// TIA Portal V20 program export: 0 tag tables, 0 data types, 16 data blocks, 79 code blocks (in call order from the OBs), 59 instance data blocks

DATA_BLOCK "Control_DB"   // DB69
{ S7_Optimized_Access := 'TRUE' }
VERSION : 0.1
// stored: AutoNumber true, DBAccessibleFromOPCUA true, DBAccessibleFromWebserver true, IsOnlyStoredInLoadMemory false, IsRetainMemResEnabled false, IsWriteProtectedInAS false, MemoryReserve 100
   VAR
      Inbound_Cnv : "Inbound_Cnv_Control_UDT";
      PopUp_Cnv { S7_SetPoint := 'True'} : Array[1..4] of "PopUp_Cnv_Control";
      Outbound_Cnv { S7_SetPoint := 'True'} : "Outbound_Cnv_Control";
      ECnv_Control { S7_SetPoint := 'True'} : "ECnv_Control";
      LCnv_Control { S7_SetPoint := 'True'} : Array[1..3] of "Buffer_Cnv_Control";
      VTD_Control { S7_SetPoint := 'True'} : "VTD_Control";
      "VTD_Order Table" { S7_SetPoint := 'True'} : "WMS_OPC_UA";
      "Carrousel_Order Table" { S7_SetPoint := 'True'} : "WMS_OPC_UA";
      Shuttles_Position : Array[1..3] of Struct
         x : DInt;
         y : DInt;
         Charging : Bool;
      END_STRUCT;
      "Weighing Station" : Struct
         Start : Bool;
         Ready : Bool;
         Running : Bool;
         Done : Bool;
         Valid : Bool;
         Weight : Real;
         Error_ID : Word;
      END_STRUCT;
      "Profiling Station" : Struct
         Start : Bool;
         Ready : Bool;
         Running : Bool;
         Done : Bool;
         Valid : Bool;
         OverWidth : Bool;
         OverHeight : Bool;
         OverLength : Bool;
         Error_ID : Word;
      END_STRUCT;
      Pick_Station : Struct
         Cnv_Occupied { ExternalWritable := 'False'} : Bool;
         PushButton : Bool;
         LightGuard : Bool;
         PushButtonLight : Bool;
         Mode { ExternalWritable := 'False'} : UInt;
         Error { ExternalWritable := 'False'} : Bool;
         Warning { ExternalWritable := 'False'} : UInt;
         Enabled { ExternalWritable := 'False'} : Bool;
         Stopped { ExternalWritable := 'False'} : Bool;
         Done : Bool;
         Running { ExternalWritable := 'False'} : Bool;
         Ready_For_Task { ExternalWritable := 'False'} : Bool;
         Current_Task_Type : UInt;
         Current_Task_ID { ExternalWritable := 'False'} : UInt;
         Pallet_Type { ExternalWritable := 'False'} : UInt;
         SM_State { ExternalWritable := 'False'} : UInt;
         Motor : "Cnv_Motor";
         Instruction : "OutCnv_Instruction";
         Cnv_Errors { S7_SetPoint := 'True'} : "Cnv_Errors";
      END_STRUCT;
      InBarcode_Station : Struct
         Start : Bool;
         Ready : Bool;
         Running : Bool;
         Done : Bool;
         Valid : Bool;
         Barcode : String;
         "Reading Gate number" : String;
         "Reading Gate number OLD" : String;
         "Number of Reading Gates" : String;
         "Number of Reading Gates OLD" : String;
      END_STRUCT;
      OutBarcode_Station : Struct
         Start : Bool;
         Ready : Bool;
         Running : Bool;
         Done : Bool;
         Valid : Bool;
         Barcode : String;
         Barcode_Old : Array[1..16] of Char;
      END_STRUCT;
      VTDBarcode_Station : Struct
         Start : Bool;
         Ready : Bool;
         Running : Bool;
         Done : Bool;
         Valid : Bool;
         Barcode : String;
         Barcode_Old : String;
      END_STRUCT;
      Movement_Completed : Struct
         RTR_ITP1 : Bool;
         RTR_P1TP2 : Bool;
         RTR_P2TP3 : Bool;
         RTR_P3TP4 : Bool;
         RTR_P4TO : Bool;
         Chain_To_Chain : Bool;
         Pop4_To_Pick : Bool;
         Pick_To_Pop1 : Bool;
         WeighingStation : Bool;
      END_STRUCT;
   END_VAR
BEGIN
END_DATA_BLOCK

DATA_BLOCK "DB_SICK_AFx60_Data"   // DB120
{ S7_Optimized_Access := 'TRUE' }
VERSION : 0.1
// stored: AutoNumber true, DBAccessibleFromOPCUA true, DBAccessibleFromWebserver true, IsOnlyStoredInLoadMemory false, IsRetainMemResEnabled false, IsWriteProtectedInAS false, MemoryReserve 100
   VAR
      Data { S7_SetPoint := 'True'} : "ST_SICK_AFx60";
   END_VAR
BEGIN
END_DATA_BLOCK

DATA_BLOCK "HMI_DB"   // DB21
{ S7_Optimized_Access := 'TRUE' }
VERSION : 0.1
// stored: AutoNumber true, DBAccessibleFromOPCUA true, DBAccessibleFromWebserver true, IsOnlyStoredInLoadMemory false, IsRetainMemResEnabled false, IsWriteProtectedInAS false, MemoryReserve 100
   VAR
      Reset : Bool;
      ChargeData : Bool;
      Username : String := 'admin';
      Password : String := '12345';
      ScreenNo : UInt;
      GeneralErrors : Word;
   END_VAR
BEGIN
END_DATA_BLOCK

DATA_BLOCK "HMI_OrderTable"   // DB110
{ S7_Optimized_Access := 'TRUE' }
VERSION : 0.1
// stored: AutoNumber true, DBAccessibleFromOPCUA true, DBAccessibleFromWebserver true, IsOnlyStoredInLoadMemory false, IsRetainMemResEnabled false, IsWriteProtectedInAS false, MemoryReserve 100
   VAR
      OrderTable_1 : Array[0..9] of "OrderTable_UDT";
      OrderTable_2 : Array[0..9] of "OrderTable_UDT";
      State_1 { S7_SetPoint := 'True'} : Array[0..9] of USInt;
      State_2 { S7_SetPoint := 'True'} : Array[0..9] of USInt;
      Index_1 : Array[0..9] of Int;
      Index_2 : Array[0..9] of Int;
      ScrollUp_PB : Bool;
      ScrollDown_PB : Bool;
      PlaceOrder_PB : Bool;
      PauseOrders_PB : Bool;
      ResumeOrder_PB : Bool;
      CancelOrder_PB : Bool;
      CancelThisOrder_PB : Bool;
      StartRow : Int;
      Device : USInt;
      PlacingNewOrder : Bool;
      PopUp_ErrorWindow_Active : Bool;
      PopUp_ErrorID : UInt;
      PopUp_Index : Int;
   END_VAR
BEGIN
END_DATA_BLOCK

DATA_BLOCK "HMI_Systems"   // DB137
{ S7_Optimized_Access := 'TRUE' }
VERSION : 0.1
// stored: AutoNumber true, DBAccessibleFromOPCUA true, DBAccessibleFromWebserver true, IsOnlyStoredInLoadMemory false, IsRetainMemResEnabled false, IsWriteProtectedInAS false, MemoryReserve 100
   VAR
      SystemNo : USInt := 1;   // System Number (1 or 2)
      System { ExternalWritable := 'False'} : "System_UDT";
      CarMeasurement { ExternalWritable := 'False'} : "CarMeasurement_DB_UDT";
      EntryGate : Struct
         Sts_Opened : Bool := TRUE;
         Sts_Closed : Bool := FALSE;
         Cmd_Open : Bool := FALSE;
         Cmd_Close : Bool := FALSE;
      END_STRUCT;
      ExitGate : Struct
         Sts_Opened : Bool := TRUE;
         Sts_Closed : Bool := FALSE;
         Cmd_Open : Bool := FALSE;
         Cmd_Close : Bool := FALSE;
      END_STRUCT;
      FieldSensors : DWord := 16#04A3_7FF3;   // Field Values of Sensors
      PanelSensors : DWord := 16#04A3_7FF3;   // Sensors to show on HMI screen
      Motors : DWord := 16#0E00_6001;   // Motors to show on HMI screen
      HMI_E_Stop_System_1 : Bool := FALSE;   // HMI Emergancy Stop Push Button for System #1
      HMI_E_Stop_System_2 : Bool := FALSE;   // HMI Emergancy Stop Push Button for System #2
      HMI_E_Stop_System_3 : Bool := FALSE;   // HMI Emergancy Stop Push Button for System #2
      Virtual_Emergency_BT : Bool := false;   // HMI Emergency Stop Push Button for General system
   END_VAR
BEGIN
   System.CancelOrders := FALSE;
   System.PauseOrders := FALSE;
   System.ResumeOrders := FALSE;
   System.OrderSent := FALSE;
   System.CurrentOrder := 0;
   System.NextOrder := 1;
   System.OrderTable[0].OrderNo := 0;
   System.OrderTable[1..34].OrderNo := -1;
   System.OrderTable[35].OrderNo := 55;
   System.OrderTable[36].OrderNo := 54;
   System.OrderTable[37..38].OrderNo := 53;
   System.OrderTable[39..45].OrderNo := -1;
   System.OrderTable[46..47].OrderNo := 52;
   System.OrderTable[48..49].OrderNo := 51;
   System.OrderTable[50].OrderNo := -1;
   System.OrderTable[51].OrderNo := 50;
   System.OrderTable[52].OrderNo := 49;
   System.OrderTable[53..54].OrderNo := 48;
   System.OrderTable[55..56].OrderNo := 47;
   System.OrderTable[57..58].OrderNo := 46;
   System.OrderTable[59..60].OrderNo := 45;
   System.OrderTable[61..67].OrderNo := 44;
   System.OrderTable[68..72].OrderNo := 43;
   System.OrderTable[73..78].OrderNo := 42;
   System.OrderTable[79..80].OrderNo := 41;
   System.OrderTable[81..82].OrderNo := 40;
   System.OrderTable[83..89].OrderNo := 39;
   System.OrderTable[90..91].OrderNo := 38;
   System.OrderTable[92..96].OrderNo := 37;
   System.OrderTable[97..99].OrderNo := 36;
   System.OrderTable[0].StepNo := 0;
   System.OrderTable[1..34].StepNo := -1;
   System.OrderTable[35..36].StepNo := 1;
   System.OrderTable[37].StepNo := 2;
   System.OrderTable[38].StepNo := 1;
   System.OrderTable[39..45].StepNo := -1;
   System.OrderTable[46].StepNo := 2;
   System.OrderTable[47].StepNo := 1;
   System.OrderTable[48].StepNo := 2;
   System.OrderTable[49].StepNo := 1;
   System.OrderTable[50].StepNo := -1;
   System.OrderTable[51..52].StepNo := 1;
   System.OrderTable[53].StepNo := 2;
   System.OrderTable[54].StepNo := 1;
   System.OrderTable[55].StepNo := 2;
   System.OrderTable[56].StepNo := 1;
   System.OrderTable[57].StepNo := 2;
   System.OrderTable[58].StepNo := 1;
   System.OrderTable[59].StepNo := 2;
   System.OrderTable[60].StepNo := 1;
   System.OrderTable[61].StepNo := 7;
   System.OrderTable[62].StepNo := 6;
   System.OrderTable[63].StepNo := 5;
   System.OrderTable[64].StepNo := 4;
   System.OrderTable[65].StepNo := 3;
   System.OrderTable[66].StepNo := 2;
   System.OrderTable[67].StepNo := 1;
   System.OrderTable[68].StepNo := 5;
   System.OrderTable[69].StepNo := 4;
   System.OrderTable[70].StepNo := 3;
   System.OrderTable[71].StepNo := 2;
   System.OrderTable[72].StepNo := 1;
   System.OrderTable[73].StepNo := 6;
   System.OrderTable[74].StepNo := 5;
   System.OrderTable[75].StepNo := 4;
   System.OrderTable[76].StepNo := 3;
   System.OrderTable[77].StepNo := 2;
   System.OrderTable[78].StepNo := 1;
   System.OrderTable[79].StepNo := 2;
   System.OrderTable[80].StepNo := 1;
   System.OrderTable[81].StepNo := 2;
   System.OrderTable[82].StepNo := 1;
   System.OrderTable[83].StepNo := 7;
   System.OrderTable[84].StepNo := 6;
   System.OrderTable[85].StepNo := 5;
   System.OrderTable[86].StepNo := 4;
   System.OrderTable[87].StepNo := 3;
   System.OrderTable[88].StepNo := 2;
   System.OrderTable[89].StepNo := 1;
   System.OrderTable[90].StepNo := 2;
   System.OrderTable[91].StepNo := 1;
   System.OrderTable[92].StepNo := 5;
   System.OrderTable[93].StepNo := 4;
   System.OrderTable[94].StepNo := 3;
   System.OrderTable[95].StepNo := 2;
   System.OrderTable[96].StepNo := 1;
   System.OrderTable[97].StepNo := 6;
   System.OrderTable[98].StepNo := 5;
   System.OrderTable[99].StepNo := 4;
   System.OrderTable[0].PlaceTime := '';
   System.OrderTable[1].PlaceTime := '06/10/2022 08:58:28';
   System.OrderTable[2].PlaceTime := '06/10/2022 08:58:01';
   System.OrderTable[3].PlaceTime := '06/10/2022 08:57:38';
   System.OrderTable[4].PlaceTime := '06/10/2022 08:56:58';
   System.OrderTable[5].PlaceTime := '06/10/2022 08:46:55';
   System.OrderTable[6].PlaceTime := '06/10/2022 08:46:40';
   System.OrderTable[7].PlaceTime := '06/10/2022 08:46:00';
   System.OrderTable[8].PlaceTime := '06/10/2022 08:45:39';
   System.OrderTable[9].PlaceTime := '06/10/2022 08:45:25';
   System.OrderTable[10].PlaceTime := '06/10/2022 08:45:12';
   System.OrderTable[11].PlaceTime := '06/10/2022 08:44:47';
   System.OrderTable[12].PlaceTime := '06/10/2022 08:44:29';
   System.OrderTable[13].PlaceTime := '06/10/2022 08:44:13';
   System.OrderTable[14].PlaceTime := '06/10/2022 08:43:18';
   System.OrderTable[15].PlaceTime := '06/10/2022 08:42:58';
   System.OrderTable[16].PlaceTime := '06/10/2022 08:41:58';
   System.OrderTable[17].PlaceTime := '06/10/2022 08:41:36';
   System.OrderTable[18].PlaceTime := '06/10/2022 08:37:44';
   System.OrderTable[19].PlaceTime := '06/10/2022 08:37:27';
   System.OrderTable[20].PlaceTime := '06/10/2022 08:37:06';
   System.OrderTable[21].PlaceTime := '06/10/2022 08:35:40';
   System.OrderTable[22].PlaceTime := '06/10/2022 08:14:06';
   System.OrderTable[23].PlaceTime := '06/10/2022 08:13:36';
   System.OrderTable[24].PlaceTime := '06/10/2022 08:09:48';
   System.OrderTable[25].PlaceTime := '06/10/2022 08:09:26';
   System.OrderTable[26].PlaceTime := '06/10/2022 08:08:29';
   System.OrderTable[27].PlaceTime := '06/10/2022 08:05:42';
   System.OrderTable[28].PlaceTime := '06/10/2022 08:04:48';
   System.OrderTable[29].PlaceTime := '06/10/2022 08:03:07';
   System.OrderTable[30].PlaceTime := '06/10/2022 08:01:46';
   System.OrderTable[31].PlaceTime := '06/10/2022 08:00:57';
   System.OrderTable[32].PlaceTime := '06/10/2022 07:54:12';
   System.OrderTable[33].PlaceTime := '06/10/2022 07:53:12';
   System.OrderTable[34].PlaceTime := '06/10/2022 07:52:34';
   System.OrderTable[35].PlaceTime := '06/09/2022 15:57:28';
   System.OrderTable[36].PlaceTime := '06/09/2022 15:54:31';
   System.OrderTable[37..38].PlaceTime := '06/09/2022 15:46:22';
   System.OrderTable[39].PlaceTime := '06/09/2022 15:44:20';
   System.OrderTable[40].PlaceTime := '06/09/2022 15:44:17';
   System.OrderTable[41].PlaceTime := '06/09/2022 15:44:09';
   System.OrderTable[42].PlaceTime := '06/09/2022 15:44:07';
   System.OrderTable[43].PlaceTime := '06/09/2022 15:42:09';
   System.OrderTable[44].PlaceTime := '06/09/2022 15:42:06';
   System.OrderTable[45].PlaceTime := '06/09/2022 15:40:52';
   System.OrderTable[46..47].PlaceTime := '06/09/2022 15:38:33';
   System.OrderTable[48..49].PlaceTime := '06/09/2022 15:37:29';
   System.OrderTable[50].PlaceTime := '06/09/2022 15:28:39';
   System.OrderTable[51].PlaceTime := '06/09/2022 15:19:41';
   System.OrderTable[52].PlaceTime := '06/09/2022 15:18:44';
   System.OrderTable[53..54].PlaceTime := '06/09/2022 15:12:55';
   System.OrderTable[55..56].PlaceTime := '06/09/2022 15:06:17';
   System.OrderTable[57..58].PlaceTime := '06/09/2022 14:58:49';
   System.OrderTable[59..60].PlaceTime := '06/09/2022 14:54:55';
   System.OrderTable[61..67].PlaceTime := '06/09/2022 14:52:23';
   System.OrderTable[68..72].PlaceTime := '06/09/2022 14:50:30';
   System.OrderTable[73..78].PlaceTime := '06/09/2022 14:49:30';
   System.OrderTable[79..80].PlaceTime := '06/09/2022 14:48:13';
   System.OrderTable[81..82].PlaceTime := '06/09/2022 14:46:58';
   System.OrderTable[83..89].PlaceTime := '06/09/2022 14:44:25';
   System.OrderTable[90..91].PlaceTime := '06/09/2022 14:37:37';
   System.OrderTable[92..96].PlaceTime := '06/09/2022 14:34:13';
   System.OrderTable[97..99].PlaceTime := '06/09/2022 14:32:56';
   System.OrderTable[0].Device := '';
   System.OrderTable[1].Device := 'TurnTable';
   System.OrderTable[2].Device := 'Dolly';
   System.OrderTable[3].Device := 'TurnTable';
   System.OrderTable[4].Device := 'Dolly';
   System.OrderTable[5..36].Device := 'Shuttle';
   System.OrderTable[37].Device := 'Dolly';
   System.OrderTable[38].Device := 'Shuttle';
   System.OrderTable[39].Device := 'Dolly';
   System.OrderTable[40].Device := 'Shuttle';
   System.OrderTable[41].Device := 'Dolly';
   System.OrderTable[42].Device := 'Shuttle';
   System.OrderTable[43].Device := 'Dolly';
   System.OrderTable[44].Device := 'Shuttle';
   System.OrderTable[45..46].Device := 'Dolly';
   System.OrderTable[47].Device := 'Shuttle';
   System.OrderTable[48].Device := 'Dolly';
   System.OrderTable[49].Device := 'Shuttle';
   System.OrderTable[50].Device := 'LoadingBay Exit';
   System.OrderTable[51..52].Device := 'Shuttle';
   System.OrderTable[53].Device := 'LoadingBay Entry';
   System.OrderTable[54].Device := 'VRC';
   System.OrderTable[55].Device := 'LoadingBay Entry';
   System.OrderTable[56].Device := 'VRC';
   System.OrderTable[57].Device := 'LoadingBay Entry';
   System.OrderTable[58].Device := 'VRC';
   System.OrderTable[59].Device := 'LoadingBay Exit';
   System.OrderTable[60..61].Device := 'VRC';
   System.OrderTable[62].Device := 'Shuttle';
   System.OrderTable[63].Device := 'Dolly';
   System.OrderTable[64].Device := 'Shuttle';
   System.OrderTable[65].Device := 'Dolly';
   System.OrderTable[66].Device := 'Shuttle';
   System.OrderTable[67].Device := 'VRC';
   System.OrderTable[68].Device := 'Shuttle';
   System.OrderTable[69].Device := 'Dolly';
   System.OrderTable[70].Device := 'TurnTable';
   System.OrderTable[71].Device := 'Shuttle';
   System.OrderTable[72].Device := 'VRC';
   System.OrderTable[73].Device := 'Dolly';
   System.OrderTable[74].Device := 'CarMeasurement';
   System.OrderTable[75].Device := 'Shuttle';
   System.OrderTable[76].Device := 'TurnTable';
   System.OrderTable[77].Device := 'Shuttle';
   System.OrderTable[78].Device := 'VRC';
   System.OrderTable[79].Device := 'LoadingBay Entry';
   System.OrderTable[80].Device := 'VRC';
   System.OrderTable[81].Device := 'LoadingBay Exit';
   System.OrderTable[82..83].Device := 'VRC';
   System.OrderTable[84].Device := 'Shuttle';
   System.OrderTable[85].Device := 'Dolly';
   System.OrderTable[86].Device := 'Shuttle';
   System.OrderTable[87].Device := 'Dolly';
   System.OrderTable[88].Device := 'Shuttle';
   System.OrderTable[89].Device := 'VRC';
   System.OrderTable[90].Device := 'LoadingBay Entry';
   System.OrderTable[91].Device := 'VRC';
   System.OrderTable[92].Device := 'Shuttle';
   System.OrderTable[93].Device := 'Dolly';
   System.OrderTable[94].Device := 'TurnTable';
   System.OrderTable[95].Device := 'Shuttle';
   System.OrderTable[96].Device := 'VRC';
   System.OrderTable[97].Device := 'Dolly';
   System.OrderTable[98].Device := 'CarMeasurement';
   System.OrderTable[99].Device := 'Shuttle';
   System.OrderTable[0].Sequence := 0;
   System.OrderTable[1..61].Sequence := 1;
   System.OrderTable[62].Sequence := 0;
   System.OrderTable[63..66].Sequence := 1;
   System.OrderTable[67].Sequence := 0;
   System.OrderTable[68..71].Sequence := 1;
   System.OrderTable[72].Sequence := 0;
   System.OrderTable[73].Sequence := 1;
   System.OrderTable[74].Sequence := 0;
   System.OrderTable[75..77].Sequence := 1;
   System.OrderTable[78].Sequence := 0;
   System.OrderTable[79..83].Sequence := 1;
   System.OrderTable[84].Sequence := 0;
   System.OrderTable[85..88].Sequence := 1;
   System.OrderTable[89].Sequence := 0;
   System.OrderTable[90..95].Sequence := 1;
   System.OrderTable[96].Sequence := 0;
   System.OrderTable[97].Sequence := 1;
   System.OrderTable[98].Sequence := 0;
   System.OrderTable[99].Sequence := 1;
   System.OrderTable[0].Status := 'Error';
   System.OrderTable[1].Status := 'Completed';
   System.OrderTable[2].Status := 'Error\Cancel';
   System.OrderTable[3].Status := 'Completed';
   System.OrderTable[4].Status := 'Error\Cancel';
   System.OrderTable[5..6].Status := 'Completed';
   System.OrderTable[7].Status := 'Canceled';
   System.OrderTable[8..10].Status := 'Completed';
   System.OrderTable[11].Status := 'Canceled';
   System.OrderTable[12..15].Status := 'Completed';
   System.OrderTable[16].Status := 'Canceled';
   System.OrderTable[17..26].Status := 'Completed';
   System.OrderTable[27].Status := 'Error\Cancel';
   System.OrderTable[28..34].Status := 'Canceled';
   System.OrderTable[35..36].Status := 'Completed';
   System.OrderTable[37].Status := 'Error\Cancel';
   System.OrderTable[38..52].Status := 'Completed';
   System.OrderTable[53].Status := 'Car Refused';
   System.OrderTable[54].Status := 'Completed';
   System.OrderTable[55].Status := 'Car Refused';
   System.OrderTable[56].Status := 'Completed';
   System.OrderTable[57].Status := 'Car Refused';
   System.OrderTable[58..89].Status := 'Completed';
   System.OrderTable[90].Status := 'Car Refused';
   System.OrderTable[91..99].Status := 'Completed';
   System.OrderTable[0].CompleteTime := '06/10/2022 08:58:15';
   System.OrderTable[1].CompleteTime := '06/10/2022 08:58:44';
   System.OrderTable[2].CompleteTime := '06/10/2022 08:58:07';
   System.OrderTable[3].CompleteTime := '06/10/2022 08:57:53';
   System.OrderTable[4].CompleteTime := '06/10/2022 08:57:03';
   System.OrderTable[5].CompleteTime := '06/10/2022 08:47:08';
   System.OrderTable[6].CompleteTime := '06/10/2022 08:46:55';
   System.OrderTable[7].CompleteTime := '06/10/2022 08:46:14';
   System.OrderTable[8].CompleteTime := '06/10/2022 08:45:52';
   System.OrderTable[9].CompleteTime := '06/10/2022 08:45:38';
   System.OrderTable[10].CompleteTime := '06/10/2022 08:45:24';
   System.OrderTable[11].CompleteTime := '06/10/2022 08:44:59';
   System.OrderTable[12].CompleteTime := '06/10/2022 08:44:41';
   System.OrderTable[13].CompleteTime := '06/10/2022 08:44:28';
   System.OrderTable[14].CompleteTime := '06/10/2022 08:43:58';
   System.OrderTable[15].CompleteTime := '06/10/2022 08:43:13';
   System.OrderTable[16].CompleteTime := '06/10/2022 08:42:28';
   System.OrderTable[17].CompleteTime := '06/10/2022 08:41:49';
   System.OrderTable[18].CompleteTime := '06/10/2022 08:37:57';
   System.OrderTable[19].CompleteTime := '06/10/2022 08:37:43';
   System.OrderTable[20].CompleteTime := '06/10/2022 08:37:19';
   System.OrderTable[21].CompleteTime := '06/10/2022 08:35:45';
   System.OrderTable[22].CompleteTime := '06/10/2022 08:14:19';
   System.OrderTable[23].CompleteTime := '06/10/2022 08:13:51';
   System.OrderTable[24].CompleteTime := '06/10/2022 08:10:02';
   System.OrderTable[25].CompleteTime := '06/10/2022 08:09:37';
   System.OrderTable[26].CompleteTime := '06/10/2022 08:08:43';
   System.OrderTable[27].CompleteTime := '06/10/2022 08:07:08';
   System.OrderTable[28].CompleteTime := '06/10/2022 08:05:11';
   System.OrderTable[29].CompleteTime := '06/10/2022 08:03:33';
   System.OrderTable[30].CompleteTime := '06/10/2022 08:02:26';
   System.OrderTable[31].CompleteTime := '06/10/2022 08:01:19';
   System.OrderTable[32].CompleteTime := '06/10/2022 08:00:14';
   System.OrderTable[33].CompleteTime := '06/10/2022 07:53:22';
   System.OrderTable[34].CompleteTime := '06/10/2022 07:52:39';
   System.OrderTable[35].CompleteTime := '06/09/2022 15:57:54';
   System.OrderTable[36].CompleteTime := '06/09/2022 15:54:58';
   System.OrderTable[37].CompleteTime := '06/09/2022 15:49:19';
   System.OrderTable[38].CompleteTime := '06/09/2022 15:46:22';
   System.OrderTable[39].CompleteTime := '06/09/2022 15:45:38';
   System.OrderTable[40].CompleteTime := '06/09/2022 15:45:09';
   System.OrderTable[41].CompleteTime := '06/09/2022 15:44:52';
   System.OrderTable[42].CompleteTime := '06/09/2022 15:44:23';
   System.OrderTable[43].CompleteTime := '06/09/2022 15:42:52';
   System.OrderTable[44].CompleteTime := '06/09/2022 15:42:22';
   System.OrderTable[45].CompleteTime := '06/09/2022 15:41:22';
   System.OrderTable[46].CompleteTime := '06/09/2022 15:39:25';
   System.OrderTable[47].CompleteTime := '06/09/2022 15:38:42';
   System.OrderTable[48].CompleteTime := '06/09/2022 15:38:27';
   System.OrderTable[49].CompleteTime := '06/09/2022 15:37:44';
   System.OrderTable[50].CompleteTime := '06/09/2022 15:28:55';
   System.OrderTable[51].CompleteTime := '06/09/2022 15:19:58';
   System.OrderTable[52].CompleteTime := '06/09/2022 15:19:11';
   System.OrderTable[53].CompleteTime := '06/09/2022 15:14:08';
   System.OrderTable[54].CompleteTime := '06/09/2022 15:12:51';
   System.OrderTable[55].CompleteTime := '06/09/2022 15:07:30';
   System.OrderTable[56].CompleteTime := '06/09/2022 15:06:13';
   System.OrderTable[57].CompleteTime := '06/09/2022 15:00:22';
   System.OrderTable[58].CompleteTime := '06/09/2022 14:58:46';
   System.OrderTable[59].CompleteTime := '06/09/2022 14:56:06';
   System.OrderTable[60].CompleteTime := '06/09/2022 14:54:51';
   System.OrderTable[61].CompleteTime := '06/09/2022 14:54:47';
   System.OrderTable[62].CompleteTime := '06/09/2022 14:54:37';
   System.OrderTable[63].CompleteTime := '06/09/2022 14:54:24';
   System.OrderTable[64].CompleteTime := '06/09/2022 14:53:55';
   System.OrderTable[65].CompleteTime := '06/09/2022 14:53:33';
   System.OrderTable[66].CompleteTime := '06/09/2022 14:52:37';
   System.OrderTable[67].CompleteTime := '06/09/2022 14:52:41';
   System.OrderTable[68].CompleteTime := '06/09/2022 14:52:18';
   System.OrderTable[69].CompleteTime := '06/09/2022 14:52:00';
   System.OrderTable[70].CompleteTime := '06/09/2022 14:51:04';
   System.OrderTable[71].CompleteTime := '06/09/2022 14:50:48';
   System.OrderTable[72].CompleteTime := '06/09/2022 14:50:49';
   System.OrderTable[73].CompleteTime := '06/09/2022 14:50:25';
   System.OrderTable[74..75].CompleteTime := '06/09/2022 14:49:55';
   System.OrderTable[76].CompleteTime := '06/09/2022 14:49:43';
   System.OrderTable[77].CompleteTime := '06/09/2022 14:49:27';
   System.OrderTable[78].CompleteTime := '06/09/2022 14:49:48';
   System.OrderTable[79].CompleteTime := '06/09/2022 14:49:23';
   System.OrderTable[80].CompleteTime := '06/09/2022 14:48:10';
   System.OrderTable[81].CompleteTime := '06/09/2022 14:47:39';
   System.OrderTable[82].CompleteTime := '06/09/2022 14:46:54';
   System.OrderTable[83].CompleteTime := '06/09/2022 14:46:50';
   System.OrderTable[84].CompleteTime := '06/09/2022 14:46:41';
   System.OrderTable[85].CompleteTime := '06/09/2022 14:46:28';
   System.OrderTable[86].CompleteTime := '06/09/2022 14:45:58';
   System.OrderTable[87].CompleteTime := '06/09/2022 14:45:37';
   System.OrderTable[88].CompleteTime := '06/09/2022 14:44:40';
   System.OrderTable[89].CompleteTime := '06/09/2022 14:44:44';
   System.OrderTable[90].CompleteTime := '06/09/2022 14:38:50';
   System.OrderTable[91].CompleteTime := '06/09/2022 14:37:33';
   System.OrderTable[92].CompleteTime := '06/09/2022 14:36:02';
   System.OrderTable[93].CompleteTime := '06/09/2022 14:35:43';
   System.OrderTable[94].CompleteTime := '06/09/2022 14:34:46';
   System.OrderTable[95].CompleteTime := '06/09/2022 14:34:31';
   System.OrderTable[96].CompleteTime := '06/09/2022 14:34:32';
   System.OrderTable[97].CompleteTime := '06/09/2022 14:34:07';
   System.OrderTable[98..99].CompleteTime := '06/09/2022 14:33:36';
   System.OrderTable[0].ErrorID := 1121;
   System.OrderTable[1].ErrorID := 0;
   System.OrderTable[2].ErrorID := 1121;
   System.OrderTable[3].ErrorID := 0;
   System.OrderTable[4].ErrorID := 1117;
   System.OrderTable[5..13].ErrorID := 0;
   System.OrderTable[14].ErrorID := 2101;
   System.OrderTable[15..26].ErrorID := 0;
   System.OrderTable[27].ErrorID := 2101;
   System.OrderTable[28..31].ErrorID := 0;
   System.OrderTable[32].ErrorID := 2104;
   System.OrderTable[33..36].ErrorID := 0;
   System.OrderTable[37].ErrorID := 1118;
   System.OrderTable[38..99].ErrorID := 0;
   System.StepTable[1..20].OrderNo := 0;
   System.StepTable[1..20].StepNo := 0;
   System.StepTable[1..20].PlaceTime := '';
   System.StepTable[1..20].Device := '';
   System.StepTable[1..20].Sequence := 0;
   System.StepTable[1..20].Status := '';
   System.StepTable[1..20].CompleteTime := '';
   System.StepTable[1..20].ErrorID := 0;
   System.CarParked_Confirm := FALSE;
   System.Running := FALSE;
   System.IDLE := TRUE;
   System.Error := FALSE;
   System.State := 0;
   System.ResetError := FALSE;
   System.Ready := TRUE;
   System.Selected := TRUE;
   System.Auto_Man := TRUE;
   System.Paused := FALSE;
   CarMeasurement.Enable := TRUE;
   CarMeasurement.Execute := FALSE;
   CarMeasurement.Cancel := FALSE;
   CarMeasurement.Enabled := TRUE;
   CarMeasurement.Done := FALSE;
   CarMeasurement.Running := FALSE;
   CarMeasurement.CarSize := 0;
   CarMeasurement.strState := 'IDLE MODE';
END_DATA_BLOCK

DATA_BLOCK "PopUps_DB"   // DB20
{ S7_Optimized_Access := 'TRUE' }
VERSION : 0.1
// stored: AutoNumber true, DBAccessibleFromOPCUA true, DBAccessibleFromWebserver true, IsOnlyStoredInLoadMemory false, IsRetainMemResEnabled false, IsWriteProtectedInAS false, MemoryReserve 100
   VAR
      Cnv_Select : DInt;
      Cnv_Select_Old : DInt;
      VTD_Select : DInt;
      Buffer_Cnv_Settings : "Buffer_Cnv_Settings";
      ECnv_Settings { S7_SetPoint := 'True'} : "ECnv_Settings";
      Inbound_Cnv_Settings { S7_SetPoint := 'True'} : "Inbound_Cnv_Settings";
      Outbound_Cnv_Settings { S7_SetPoint := 'True'} : "Outbound_Cnv_Settings";
      PopUp_Cnv_settings { S7_SetPoint := 'True'} : "PopUp_Cnv_Settings";
      System_Settings { S7_SetPoint := 'True'} : "System_Settings";
      VTD_Settings { S7_SetPoint := 'True'} : "VTD_Settings";
      Shuttle_MQTT_Settings { S7_SetPoint := 'True'} : "MQTT_Settings";
      LockingPins : Struct
         Faceplate : "FacePlate_LP_UDT";
         ExtendLeft { S7_SetPoint := 'True'} : Bool;
         RetractLeft { S7_SetPoint := 'True'} : Bool;
         ExtendRight { S7_SetPoint := 'True'} : Bool;
         RetractRight { S7_SetPoint := 'True'} : Bool;
         Extend_All : Bool;
         Retract_All : Bool;
      END_STRUCT;
      BSettings_Visibility : Bool;
      ESettings_Visibility : Bool;
      InSettings_Visibility : Bool;
      OutSettings_Visibility : Bool;
      PSettings_Visibility : Bool;
   END_VAR
BEGIN
   Shuttle_MQTT_Settings.MQTT_Con_Params.hwId := 64;
   Shuttle_MQTT_Settings.MQTT_Con_Params.broker := '10.0.34.2';
   Shuttle_MQTT_Settings.Client_ID := WSTRING#'PLC';
   Shuttle_MQTT_Settings.Username := WSTRING#'Devin';
   Shuttle_MQTT_Settings.Password := WSTRING#'1';
   Shuttle_MQTT_Settings.Retain := TRUE;
END_DATA_BLOCK

DATA_BLOCK "SAI_Buffer"   // DB600
{ S7_Optimized_Access := 'FALSE' }
VERSION : 0.1
// stored: AutoNumber false, DBAccessibleFromOPCUA true, DBAccessibleFromWebserver true, IsOnlyStoredInLoadMemory false, IsWriteProtectedInAS false
   VAR RETAIN
      WriteBuf : Array[0..3] of Byte;
      ReadBuf : Array[0..3] of Byte;
   END_VAR
BEGIN
END_DATA_BLOCK

DATA_BLOCK "SAI_IND_AlibiData"   // DB106
{ S7_Optimized_Access := 'TRUE' }
VERSION : 0.1
// stored: AutoNumber true, DBAccessibleFromOPCUA true, DBAccessibleFromWebserver true, IsOnlyStoredInLoadMemory false, IsRetainMemResEnabled false, IsWriteProtectedInAS false, MemoryReserve 100
   VAR
      Alibi_RawData : Array[0..44] of Byte;
   END_VAR
BEGIN
END_DATA_BLOCK

DATA_BLOCK "SICK_Lector"   // DB46
{ S7_Optimized_Access := 'TRUE' }
VERSION : 0.1
// stored: AutoNumber true, DBAccessibleFromOPCUA true, DBAccessibleFromWebserver true, IsOnlyStoredInLoadMemory false, IsRetainMemResEnabled false, IsWriteProtectedInAS false, MemoryReserve 100
   VAR
      Barcode_Result : String;
      HWInputIdent : HW_IO := 554;
      HWInputLength : USInt := 32;
      HWOutputIdent : HW_IO := 555;
      HWOutputLength : USInt := 32;
      CANId : USInt := 0;
      TOut : Time := T#10S;
      Req : Bool := FALSE;
      TriggerOn : Bool := FALSE;
      TriggerOff : Bool := FALSE;
      Matchcode : Bool := FALSE;
      SavePermanent : Bool := FALSE;
      ComTest : Bool := FALSE;
      FreeCommand : Bool := FALSE;
      Data : "ST_SICK_Lector_CLV6xx";
      RdDone { S7_SetPoint := 'True'} : Bool := FALSE;
      ReqDone : Bool := FALSE;
      ReqBusy : Bool := FALSE;
      Error : Bool := TRUE;
      Errorcode : DWord := 16#0000_0015;
   END_VAR
BEGIN
   Data.Matchcode.sName := '';
   Data.Matchcode.nCodeType := ' ';
   Data.Matchcode.iMinMaxLength := 0;
   Data.Matchcode.sContent := '';
   Data.FreeCommand.sCommand := '';
   Data.FreeCommand.sResult := '';
   Data.ReadingResult.iCounter := 0;
   Data.ReadingResult.iLength := 0;
   Data.ReadingResult.arrResult[1..200] := 16#00;
END_DATA_BLOCK

DATA_BLOCK "Screen_DB"   // DB23
{ S7_Optimized_Access := 'TRUE' }
VERSION : 0.1
// stored: AutoNumber true, DBAccessibleFromOPCUA true, DBAccessibleFromWebserver true, IsOnlyStoredInLoadMemory false, IsRetainMemResEnabled false, IsWriteProtectedInAS false, MemoryReserve 100
   VAR
      VTD_LevelDetect { S7_SetPoint := 'True'} : Array[1..8] of Bool;
      VTD_Semi_CMD : Array[1..8] of Bool;
      VTD_ActualPosition { S7_SetPoint := 'True'} : DInt;
      VTD_OvertravelUp : Bool;
      VTD_LimitUp : Bool;
      VTD_CreepUp : Bool;
      VTD_SlowDownUp : Bool;
      VTD_SlowDownDown : Bool;
      VTD_CreepDown : Bool;
      VTD_LimitDown : Bool;
      VTD_OvertravelDown : Bool;
      VTD_LiftUp : Bool;
      VTD_LiftDown : Bool;
      VTD_LimitOverride : Bool;
      VTD_Manual : Bool;
      VTD_Semi : Bool;
      VTD_MemoryLatch : Bool;
      VTD_SaveData : Bool;
      VTD_Select : USInt;
      Cnv_Manual : Bool;
      Cnv_Semi : Bool;
      Cnv_Foward : Bool;
      Cnv_Backward : Bool;
      Cnv_LeftAllign : Bool;
      Cnv_RightAllign : Bool;
      Cnv_FowardTransfer : Bool;
      Cnv_BackwardTransfer : Bool;
      Cnv_ShuttleStopper : Bool;
      Cnv_ShuttleStopperVisibility : Bool;
      Cnv_Plallet_Type1Visibility : Bool;
      Cnv_Plallet_Type2Visibility : Bool;
      Cnv_Select : USInt;
      Shuttle_Status : "Shuttle_MQTT_Status_Msg";
      Shuttle_Name { S7_SetPoint := 'True'} : String;
      Shuttle_URL : String;
      Settings_ActivePopUp : USInt;
      Alarms_ActiveTable : USInt;
      MainTemplate_ErrorActive : Bool;
      MainTemplate_ErrorCount : USInt;
      MainTemplate_ScreenNo : UInt;
      MainTemplate_Background : USInt;
      EmptyTemplate_Background : USInt;
      IO_ActivePopup : USInt;
      Charge_VTD : Bool;
      Charge_Cnv : Bool;
      Charge_VTD_Commands : Bool;
      Charge_Cnv_Commands : Bool;
      Shuttle : "Shuttle_MQTT_Status_Msg";
      Shuttle_Select : USInt;
   END_VAR
BEGIN
END_DATA_BLOCK

DATA_BLOCK "Settings_DB"   // DB71
{ S7_Optimized_Access := 'TRUE' }
VERSION : 0.1
// stored: AutoNumber true, DBAccessibleFromOPCUA true, DBAccessibleFromWebserver true, IsOnlyStoredInLoadMemory false, IsRetainMemResEnabled false, IsWriteProtectedInAS false, MemoryReserve 100
   VAR RETAIN
      Inbound_Cnv_Settings { S7_SetPoint := 'True'} : "Inbound_Cnv_Settings";
      PopUp_Cnv_Settings { S7_SetPoint := 'True'} : Array[1..4] of "PopUp_Cnv_Settings";
      Pick_Cnv_Settings { S7_SetPoint := 'True'} : "Pick_Cnv_Settings";
      Outbound_Cnv_Settings { S7_SetPoint := 'True'} : "Outbound_Cnv_Settings";
      VTD_Settings : "VTD_Settings";
      ECnv_Settings : "ECnv_Settings";
      LCnv_Settings : Array[1..3] of "Buffer_Cnv_Settings";
   END_VAR
   VAR
      "Weighing Station" : Struct
         "Minimum Weight" : Real := 30.0;
         "Maximum Weigh" : Real := 1500.0;
      END_STRUCT;
      "Profile Station" : Struct
         "Maximum Length" : Real := 1230.0;
         "Conveyor Speed mm_s" : Real := 10.0;
      END_STRUCT;
   END_VAR
   VAR RETAIN
      Shuttle_MQTT_Settings : "MQTT_Settings";
      System_Settings : "System_Settings";
   END_VAR
   VAR
      TimeStartBoost_P2ToP3 { S7_SetPoint := 'True'} : UInt := 20;
      TimeStartBoost_P3ToP4 : UInt := 8;
      TimeStartBoost_P1ToP2 : UInt := 8;
   END_VAR
BEGIN
   Inbound_Cnv_Settings.ID := 130001;
   Inbound_Cnv_Settings.TC_Time := 0;
   Inbound_Cnv_Settings.Transfer_Time := 30;
   Inbound_Cnv_Settings.Slow_Speed := 0;
   Inbound_Cnv_Settings.Full_Speed := 60;
   Inbound_Cnv_Settings.Manual_Speed := 60;
   Inbound_Cnv_Settings.No_Forklift_Detect_Timer := 5;
   Inbound_Cnv_Settings.G120_Hardware_ID := 376;
   PopUp_Cnv_Settings[1].ID := 150001;
   PopUp_Cnv_Settings[2].ID := 160001;
   PopUp_Cnv_Settings[3].ID := 170001;
   PopUp_Cnv_Settings[4].ID := 180001;
   PopUp_Cnv_Settings[1..4].Roller_TC_Time := 0;
   PopUp_Cnv_Settings[1..2].Roller_Transfer_Time := 30;
   PopUp_Cnv_Settings[3..4].Roller_Transfer_Time := 25;
   PopUp_Cnv_Settings[1..4].Roller_Slow_Speed := 0;
   PopUp_Cnv_Settings[1..4].Roller_Full_Speed := 60;
   PopUp_Cnv_Settings[1..3].Roller_Manual_Speed := 60;
   PopUp_Cnv_Settings[4].Roller_Manual_Speed := 50;
   PopUp_Cnv_Settings[1..4].Chain_TC_Time := 0;
   PopUp_Cnv_Settings[1].Chain_Transfer_Time := 50;
   PopUp_Cnv_Settings[2].Chain_Transfer_Time := 500;
   PopUp_Cnv_Settings[3].Chain_Transfer_Time := 40;
   PopUp_Cnv_Settings[4].Chain_Transfer_Time := 50;
   PopUp_Cnv_Settings[1..2].Chain_Slow_Speed := 0;
   PopUp_Cnv_Settings[3].Chain_Slow_Speed := 50;
   PopUp_Cnv_Settings[4].Chain_Slow_Speed := 0;
   PopUp_Cnv_Settings[1].Chain_Full_Speed := 60;
   PopUp_Cnv_Settings[2..3].Chain_Full_Speed := 70;
   PopUp_Cnv_Settings[4].Chain_Full_Speed := 60;
   PopUp_Cnv_Settings[1].Chain_Manual_Speed := 30;
   PopUp_Cnv_Settings[2].Chain_Manual_Speed := 60;
   PopUp_Cnv_Settings[3].Chain_Manual_Speed := 50;
   PopUp_Cnv_Settings[4].Chain_Manual_Speed := 60;
   PopUp_Cnv_Settings[1..4].Lift_TC_Time := 0;
   PopUp_Cnv_Settings[1].Lift_Transfer_Time := 7;
   PopUp_Cnv_Settings[2..4].Lift_Transfer_Time := 15;
   PopUp_Cnv_Settings[1..4].Lift_Slow_Speed := 0;
   PopUp_Cnv_Settings[1..2].Lift_Full_Speed := 100;
   PopUp_Cnv_Settings[3].Lift_Full_Speed := 80;
   PopUp_Cnv_Settings[4].Lift_Full_Speed := 100;
   PopUp_Cnv_Settings[1].Lift_Manual_Speed := 40;
   PopUp_Cnv_Settings[2..4].Lift_Manual_Speed := 10;
   PopUp_Cnv_Settings[1].Roller_G120_Hardware_ID := 385;
   PopUp_Cnv_Settings[2].Roller_G120_Hardware_ID := 394;
   PopUp_Cnv_Settings[3].Roller_G120_Hardware_ID := 403;
   PopUp_Cnv_Settings[4].Roller_G120_Hardware_ID := 466;
   PopUp_Cnv_Settings[1].Chain_G120_Hardware_ID := 412;
   PopUp_Cnv_Settings[2].Chain_G120_Hardware_ID := 421;
   PopUp_Cnv_Settings[3].Chain_G120_Hardware_ID := 430;
   PopUp_Cnv_Settings[4].Chain_G120_Hardware_ID := 0;
   PopUp_Cnv_Settings[1].Lift_G120_Hardware_ID := 340;
   PopUp_Cnv_Settings[2].Lift_G120_Hardware_ID := 358;
   PopUp_Cnv_Settings[3].Lift_G120_Hardware_ID := 493;
   PopUp_Cnv_Settings[4].Lift_G120_Hardware_ID := 349;
   Pick_Cnv_Settings.ID := 410001;
   Pick_Cnv_Settings.TC_Time := 0;
   Pick_Cnv_Settings.Transfer_Time := 25;
   Pick_Cnv_Settings.Slow_Speed := 0;
   Pick_Cnv_Settings.Full_Speed := 60;
   Pick_Cnv_Settings.Manual_Speed := 60;
   Pick_Cnv_Settings.No_Forklift_Detect_Timer := 0;
   Pick_Cnv_Settings.G120_Hardware_ID := 412;
   Outbound_Cnv_Settings.ID := 140001;
   Outbound_Cnv_Settings.TC_Time := 0;
   Outbound_Cnv_Settings.Transfer_Time := 25;
   Outbound_Cnv_Settings.Slow_Speed := 0;
   Outbound_Cnv_Settings.Full_Speed := 60;
   Outbound_Cnv_Settings.Manual_Speed := 60;
   Outbound_Cnv_Settings.No_Forklift_Detect_Timer := 5;
   Outbound_Cnv_Settings.G120_Hardware_ID := 367;
   VTD_Settings.ID := 1;
   VTD_Settings.Lowest_Level := 1;
   VTD_Settings.Highest_Level := 3;
   VTD_Settings.VTD_Max_Heigh := 7145;
   VTD_Settings.VTD_Min_Height := 68;
   VTD_Settings.VTD_Level_Granularity := 20;
   VTD_Settings.Dft_Level_Offset_LE := 0;
   VTD_Settings.Dft_Level_Offset_AE := 0;
   VTD_Settings.Teach_Speed := 0;
   VTD_Settings.Creep_Speed := 5;
   VTD_Settings.Slow_Speed := 5;
   VTD_Settings.Slow_Calib_Speed := 5;
   VTD_Settings.Loaded_Speed := 80;
   VTD_Settings.Shuttle_Speed := 80;
   VTD_Settings.Pallet_Speed := 40;
   VTD_Settings.Empty_Speed := 60;
   VTD_Settings.Dock_speed := 5;
   VTD_Settings.Manual_Speed := 10;
   VTD_Settings.Slowdown_Count_LE := 600;
   VTD_Settings.Creep_Count_LE := 60;
   VTD_Settings.Slowdown_Count_AE := 700;
   VTD_Settings.Creep_Count_AE := 60;
   VTD_Settings.Encoder_Delta_W1 := 0.0;
   VTD_Settings.Encoder_Delta_W2 := 0.0;
   VTD_Settings.AE_Ratio := 0.0;
   VTD_Settings.Encoder_Delta_Warning := 60.0;
   VTD_Settings.Encoder_Delta_Error := 80.0;
   VTD_Settings.Transfer_Timeout_Up := 200;
   VTD_Settings.Transfer_Timeout_Down := 200;
   VTD_Settings.Lockpins_Timeout_Extend := 6000;
   VTD_Settings.Lockpins_Timeout_Retract := 6000;
   VTD_Settings.Level_Detect_Timeout := 500;
   VTD_Settings.Teach_Timeout := 600;
   VTD_Settings.Chain_Slack_Timeout := 700;
   VTD_Settings.Level_Detect_LE := 3.0;
   VTD_Settings.G120_Hardware_ID := 612;
   VTD_Settings.Teach_Values.Levels_LE[0] := 69.0;
   VTD_Settings.Teach_Values.Levels_LE[1] := 3451.0;
   VTD_Settings.Teach_Values.Levels_LE[2] := 5249.0;
   VTD_Settings.Teach_Values.Levels_LE[3] := 7049.0;
   VTD_Settings.Teach_Values.Levels_AE[0] := 0;
   VTD_Settings.Teach_Values.Levels_AE[1] := 63;
   VTD_Settings.Teach_Values.Levels_AE[2] := 2069;
   VTD_Settings.Teach_Values.Levels_AE[3] := 4077;
   ECnv_Settings.ID := 120101;
   ECnv_Settings.Barcode_ID := 0;
   ECnv_Settings.Cnv_Level := 1;
   ECnv_Settings.TC_Time := 0;
   ECnv_Settings.Transfer_Time := 20;
   ECnv_Settings.Pallet_Align_Time := 0;
   ECnv_Settings.Slow_Speed := 0;
   ECnv_Settings.Full_Speed := 70;
   ECnv_Settings.Manual_Speed := 50;
   ECnv_Settings.G120_Hardware_ID := 475;
   LCnv_Settings[1].ID := 100101;
   LCnv_Settings[2].ID := 100201;
   LCnv_Settings[3].ID := 100301;
   LCnv_Settings[1..3].Barcode_ID := 0;
   LCnv_Settings[1].Cnv_Level := 1;
   LCnv_Settings[2].Cnv_Level := 2;
   LCnv_Settings[3].Cnv_Level := 3;
   LCnv_Settings[1..3].TC_Time := 1;
   LCnv_Settings[1..3].Transfer_Time := 20;
   LCnv_Settings[1..3].Pallet_Align_Time := 4;
   LCnv_Settings[1..3].Slow_Speed := 25;
   LCnv_Settings[1..3].Full_Speed := 70;
   LCnv_Settings[1..2].Manual_Speed := 60;
   LCnv_Settings[3].Manual_Speed := 50;
   LCnv_Settings[1..3].Safety_stop_Timeout := 0;
   LCnv_Settings[1].G120_Hardware_ID := 439;
   LCnv_Settings[2].G120_Hardware_ID := 448;
   LCnv_Settings[3].G120_Hardware_ID := 457;
   Shuttle_MQTT_Settings.MQTT_Con_Params.hwId := 64;
   Shuttle_MQTT_Settings.MQTT_Con_Params.connId := 16#0001;
   Shuttle_MQTT_Settings.MQTT_Con_Params.broker := '10.0.34.2';
   Shuttle_MQTT_Settings.MQTT_Con_Params.port := 1883;
   Shuttle_MQTT_Settings.MQTT_Con_Params.tls.enableTls := FALSE;
   Shuttle_MQTT_Settings.MQTT_Con_Params.tls.validateServerIdentity := FALSE;
   Shuttle_MQTT_Settings.MQTT_Con_Params.tls.brokerCert := 0;
   Shuttle_MQTT_Settings.MQTT_Con_Params.tls.clientCert := 0;
   Shuttle_MQTT_Settings.MQTT_Con_Params.keepAlive := 60;
   Shuttle_MQTT_Settings.Client_ID := WSTRING#'PLC';
   Shuttle_MQTT_Settings.Username := WSTRING#'Devin';
   Shuttle_MQTT_Settings.Password := WSTRING#'1';
   Shuttle_MQTT_Settings.Timeout := 0;
   Shuttle_MQTT_Settings.QoS := 0;
   Shuttle_MQTT_Settings.Retain := TRUE;
   Shuttle_MQTT_Settings.Will_Topic := WSTRING#'';
   Shuttle_MQTT_Settings.Will_Msg_Length := 0;
   Shuttle_MQTT_Settings.Will_Msg_Payload[1..128] := 16#00;
   System_Settings.VTD_Count := 1;
   System_Settings.Level_Count := 3;
   System_Settings.Cnv_Count := 10;
   System_Settings.Shuttle_Count := 3;
   System_Settings.Shuttle_Interlock_Timeout := 999;
END_DATA_BLOCK

DATA_BLOCK "Shuttle_MQTT_DB"   // DB75
{ S7_Optimized_Access := 'TRUE' }
VERSION : 0.1
// stored: AutoNumber true, DBAccessibleFromOPCUA true, DBAccessibleFromWebserver true, IsOnlyStoredInLoadMemory false, IsRetainMemResEnabled false, IsWriteProtectedInAS false, MemoryReserve 100
   VAR
      Shuttle_MQTT : Array[1..3] of "MQTT_Interface";
   END_VAR
BEGIN
END_DATA_BLOCK

DATA_BLOCK "TCP_IP_DB_Estop_Shuttle1"   // DB166
{ S7_Optimized_Access := 'TRUE' }
VERSION : 0.1
// stored: AutoNumber false, DBAccessibleFromOPCUA true, DBAccessibleFromWebserver true, IsOnlyStoredInLoadMemory false, IsRetainMemResEnabled false, IsWriteProtectedInAS false, MemoryReserve 100
   VAR
      enable : Bool := TRUE;
      send : Bool;
      sendDataLength : UDInt := 0;
      receiveDataLength : UDInt := 16#FFFF_FFFF;
   END_VAR
   VAR RETAIN
      tcpConfig : "LCom_typeConfig";
   END_VAR
   VAR
      tcpDiagnostics { S7_SetPoint := 'True'} : "LCom_typeDiagnostics";
      sendBuffer { S7_SetPoint := 'True'} : Array[0..59] of Byte;
      SendBufferSize : UInt := 60;
      receiveBuffer : Array[0..27] of Byte;
      receiveBufferSize : UInt := 28;
      connected : Bool;
      sending : Bool;
      dataReceived : Bool;
      receivedDataLength : UDInt;
      busy : Bool;
      error : Bool;
      status : Word;
   END_VAR
BEGIN
   tcpConfig.connection.interfaceID := 64;
   tcpConfig.connection.connectionID := 101;
   tcpConfig.connection.comService := 1;
   tcpConfig.connection.isClient := False;
   tcpConfig.connection.connectType := 1;
   tcpConfig.connection.localPort := 4001;
   tcpConfig.connection.partnerPort := 4001;
   tcpConfig.connection.partnerIP.ADDR[1] := 10;
   tcpConfig.connection.partnerIP.ADDR[2] := 0;
   tcpConfig.connection.partnerIP.ADDR[3] := 34;
   tcpConfig.connection.partnerIP.ADDR[4] := 180;
   tcpConfig.connection.acceptUnknownPartner := False;
   tcpConfig.connection.lifeSignCycleTime := T#1s;
   // sendBuffer[0] : STX
   // sendBuffer[1] : Size
   // sendBuffer[2] : Type
   // sendBuffer[3] : Request ID 1
   // sendBuffer[4] : Request ID 2
   // sendBuffer[5] : PID 1
   // sendBuffer[6] : PID 2
   // sendBuffer[7] : PID 3
   // sendBuffer[8] : PID 4
   // sendBuffer[9] : DID 1
   // sendBuffer[10] : DID 2
   // sendBuffer[11] : DID 3
   // sendBuffer[12] : DID 4
   // sendBuffer[13] : Distance remaining 1
   // sendBuffer[14] : Distance remaining 2
   // sendBuffer[15] : X
   // sendBuffer[16] : X
   // sendBuffer[17] : X
   // sendBuffer[18] : X
   // sendBuffer[19] : Y
   // sendBuffer[20] : Y
   // sendBuffer[21] : Y
   // sendBuffer[22] : Y
   // sendBuffer[23] : Floor
   // sendBuffer[24] : Mode
   // sendBuffer[25] : State
   // sendBuffer[26] : Load State
   // sendBuffer[27] : E1
   // sendBuffer[28] : E1
   // sendBuffer[29] : E2
   // sendBuffer[30] : E2
   // sendBuffer[31] : E3
   // sendBuffer[32] : E3
   // sendBuffer[33] : E4
   // sendBuffer[34] : E4
   // sendBuffer[35] : E5
   // sendBuffer[36] : E5
   // sendBuffer[37] : E6
   // sendBuffer[38] : E6
   // sendBuffer[39] : I1
   // sendBuffer[40] : I1
   // sendBuffer[41] : Q1
   // sendBuffer[42] : Q1
   // sendBuffer[43] : Barcode 1
   // sendBuffer[44] : Barcode 2
   // sendBuffer[45] : Barcode 3
   // sendBuffer[46] : Barcode 4
   // sendBuffer[47] : Pallet Type
   // sendBuffer[48] : Energy Level
   // sendBuffer[49] : Battery Voltage
   // sendBuffer[50] : Battery Voltage
   // sendBuffer[51] : Paused
   // sendBuffer[52] : Last order 1
   // sendBuffer[53] : Last order 2
   // sendBuffer[54] : Current order 1
   // sendBuffer[55] : Current order 2
   // sendBuffer[56] : Last finished 1
   // sendBuffer[57] : Last Finished 2
   // sendBuffer[58] : CS
   // sendBuffer[59] : ETX
   // receiveBuffer[0] : STX
   // receiveBuffer[1] : Size (length of payload)
   // receiveBuffer[2] : Type
   // receiveBuffer[3] : Request ID 1
   // receiveBuffer[4] : Request ID 2
END_DATA_BLOCK

DATA_BLOCK "TCP_IP_DB_Estop_Shuttle2"   // DB180
{ S7_Optimized_Access := 'TRUE' }
VERSION : 0.1
// stored: AutoNumber false, DBAccessibleFromOPCUA true, DBAccessibleFromWebserver true, IsOnlyStoredInLoadMemory false, IsRetainMemResEnabled false, IsWriteProtectedInAS false, MemoryReserve 100
   VAR
      enable : Bool := TRUE;
      send : Bool;
      sendDataLength : UDInt := 0;
      receiveDataLength : UDInt := 16#FFFF_FFFF;
   END_VAR
   VAR RETAIN
      tcpConfig : "LCom_typeConfig";
   END_VAR
   VAR
      tcpDiagnostics { S7_SetPoint := 'True'} : "LCom_typeDiagnostics";
      sendBuffer { S7_SetPoint := 'True'} : Array[0..59] of Byte;
      SendBufferSize : UInt := 60;
      receiveBuffer : Array[0..27] of Byte;
      receiveBufferSize : UInt := 28;
      connected : Bool;
      sending : Bool;
      dataReceived : Bool;
      receivedDataLength : UDInt;
      busy : Bool;
      error : Bool;
      status : Word;
   END_VAR
BEGIN
   tcpConfig.connection.interfaceID := 64;
   tcpConfig.connection.connectionID := 102;
   tcpConfig.connection.comService := 1;
   tcpConfig.connection.isClient := False;
   tcpConfig.connection.connectType := 1;
   tcpConfig.connection.localPort := 4002;
   tcpConfig.connection.partnerPort := 4002;
   tcpConfig.connection.partnerIP.ADDR[1] := 10;
   tcpConfig.connection.partnerIP.ADDR[2] := 0;
   tcpConfig.connection.partnerIP.ADDR[3] := 34;
   tcpConfig.connection.partnerIP.ADDR[4] := 185;
   tcpConfig.connection.acceptUnknownPartner := False;
   tcpConfig.connection.lifeSignCycleTime := T#1s;
   // sendBuffer[0] : STX
   // sendBuffer[1] : Size
   // sendBuffer[2] : Type
   // sendBuffer[3] : Request ID 1
   // sendBuffer[4] : Request ID 2
   // sendBuffer[5] : PID 1
   // sendBuffer[6] : PID 2
   // sendBuffer[7] : PID 3
   // sendBuffer[8] : PID 4
   // sendBuffer[9] : DID 1
   // sendBuffer[10] : DID 2
   // sendBuffer[11] : DID 3
   // sendBuffer[12] : DID 4
   // sendBuffer[13] : Distance remaining 1
   // sendBuffer[14] : Distance remaining 2
   // sendBuffer[15] : X
   // sendBuffer[16] : X
   // sendBuffer[17] : X
   // sendBuffer[18] : X
   // sendBuffer[19] : Y
   // sendBuffer[20] : Y
   // sendBuffer[21] : Y
   // sendBuffer[22] : Y
   // sendBuffer[23] : Floor
   // sendBuffer[24] : Mode
   // sendBuffer[25] : State
   // sendBuffer[26] : Load State
   // sendBuffer[27] : E1
   // sendBuffer[28] : E1
   // sendBuffer[29] : E2
   // sendBuffer[30] : E2
   // sendBuffer[31] : E3
   // sendBuffer[32] : E3
   // sendBuffer[33] : E4
   // sendBuffer[34] : E4
   // sendBuffer[35] : E5
   // sendBuffer[36] : E5
   // sendBuffer[37] : E6
   // sendBuffer[38] : E6
   // sendBuffer[39] : I1
   // sendBuffer[40] : I1
   // sendBuffer[41] : Q1
   // sendBuffer[42] : Q1
   // sendBuffer[43] : Barcode 1
   // sendBuffer[44] : Barcode 2
   // sendBuffer[45] : Barcode 3
   // sendBuffer[46] : Barcode 4
   // sendBuffer[47] : Pallet Type
   // sendBuffer[48] : Energy Level
   // sendBuffer[49] : Battery Voltage
   // sendBuffer[50] : Battery Voltage
   // sendBuffer[51] : Paused
   // sendBuffer[52] : Last order 1
   // sendBuffer[53] : Last order 2
   // sendBuffer[54] : Current order 1
   // sendBuffer[55] : Current order 2
   // sendBuffer[56] : Last finished 1
   // sendBuffer[57] : Last Finished 2
   // sendBuffer[58] : CS
   // sendBuffer[59] : ETX
   // receiveBuffer[0] : STX
   // receiveBuffer[1] : Size (length of payload)
   // receiveBuffer[2] : Type
   // receiveBuffer[3] : Request ID 1
   // receiveBuffer[4] : Request ID 2
END_DATA_BLOCK

DATA_BLOCK "TCP_IP_DB_Estop_Shuttle3"   // DB184
{ S7_Optimized_Access := 'TRUE' }
VERSION : 0.1
// stored: AutoNumber false, DBAccessibleFromOPCUA true, DBAccessibleFromWebserver true, IsOnlyStoredInLoadMemory false, IsRetainMemResEnabled false, IsWriteProtectedInAS false, MemoryReserve 100
   VAR
      enable : Bool := TRUE;
      send : Bool;
      sendDataLength : UDInt := 0;
      receiveDataLength : UDInt := 16#FFFF_FFFF;
   END_VAR
   VAR RETAIN
      tcpConfig : "LCom_typeConfig";
   END_VAR
   VAR
      tcpDiagnostics { S7_SetPoint := 'True'} : "LCom_typeDiagnostics";
      sendBuffer { S7_SetPoint := 'True'} : Array[0..59] of Byte;
      SendBufferSize : UInt := 60;
      receiveBuffer : Array[0..27] of Byte;
      receiveBufferSize : UInt := 28;
      connected : Bool;
      sending : Bool;
      dataReceived : Bool;
      receivedDataLength : UDInt;
      busy : Bool;
      error : Bool;
      status : Word;
   END_VAR
BEGIN
   tcpConfig.connection.interfaceID := 64;
   tcpConfig.connection.connectionID := 103;
   tcpConfig.connection.comService := 1;
   tcpConfig.connection.isClient := False;
   tcpConfig.connection.connectType := 1;
   tcpConfig.connection.localPort := 4003;
   tcpConfig.connection.partnerPort := 4003;
   tcpConfig.connection.partnerIP.ADDR[1] := 10;
   tcpConfig.connection.partnerIP.ADDR[2] := 0;
   tcpConfig.connection.partnerIP.ADDR[3] := 34;
   tcpConfig.connection.partnerIP.ADDR[4] := 190;
   tcpConfig.connection.acceptUnknownPartner := False;
   tcpConfig.connection.lifeSignCycleTime := T#1s;
   // sendBuffer[0] : STX
   // sendBuffer[1] : Size
   // sendBuffer[2] : Type
   // sendBuffer[3] : Request ID 1
   // sendBuffer[4] : Request ID 2
   // sendBuffer[5] : PID 1
   // sendBuffer[6] : PID 2
   // sendBuffer[7] : PID 3
   // sendBuffer[8] : PID 4
   // sendBuffer[9] : DID 1
   // sendBuffer[10] : DID 2
   // sendBuffer[11] : DID 3
   // sendBuffer[12] : DID 4
   // sendBuffer[13] : Distance remaining 1
   // sendBuffer[14] : Distance remaining 2
   // sendBuffer[15] : X
   // sendBuffer[16] : X
   // sendBuffer[17] : X
   // sendBuffer[18] : X
   // sendBuffer[19] : Y
   // sendBuffer[20] : Y
   // sendBuffer[21] : Y
   // sendBuffer[22] : Y
   // sendBuffer[23] : Floor
   // sendBuffer[24] : Mode
   // sendBuffer[25] : State
   // sendBuffer[26] : Load State
   // sendBuffer[27] : E1
   // sendBuffer[28] : E1
   // sendBuffer[29] : E2
   // sendBuffer[30] : E2
   // sendBuffer[31] : E3
   // sendBuffer[32] : E3
   // sendBuffer[33] : E4
   // sendBuffer[34] : E4
   // sendBuffer[35] : E5
   // sendBuffer[36] : E5
   // sendBuffer[37] : E6
   // sendBuffer[38] : E6
   // sendBuffer[39] : I1
   // sendBuffer[40] : I1
   // sendBuffer[41] : Q1
   // sendBuffer[42] : Q1
   // sendBuffer[43] : Barcode 1
   // sendBuffer[44] : Barcode 2
   // sendBuffer[45] : Barcode 3
   // sendBuffer[46] : Barcode 4
   // sendBuffer[47] : Pallet Type
   // sendBuffer[48] : Energy Level
   // sendBuffer[49] : Battery Voltage
   // sendBuffer[50] : Battery Voltage
   // sendBuffer[51] : Paused
   // sendBuffer[52] : Last order 1
   // sendBuffer[53] : Last order 2
   // sendBuffer[54] : Current order 1
   // sendBuffer[55] : Current order 2
   // sendBuffer[56] : Last finished 1
   // sendBuffer[57] : Last Finished 2
   // sendBuffer[58] : CS
   // sendBuffer[59] : ETX
   // receiveBuffer[0] : STX
   // receiveBuffer[1] : Size (length of payload)
   // receiveBuffer[2] : Type
   // receiveBuffer[3] : Request ID 1
   // receiveBuffer[4] : Request ID 2
END_DATA_BLOCK

DATA_BLOCK "Time"   // DB135
{ S7_Optimized_Access := 'TRUE' }
VERSION : 0.1
// stored: AutoNumber true, DBAccessibleFromOPCUA true, DBAccessibleFromWebserver true, IsOnlyStoredInLoadMemory false, IsRetainMemResEnabled false, IsWriteProtectedInAS false, MemoryReserve 100
   VAR
      CurrentLocalTime : String := '06/10/2022 09:04:28';
      CurrentDTL : DTL := DTL#2022-06-10-09:04:28.050899826;
      PC_HeartBeat : Word := 16#6E87;
      PLC_HeartBeat : Word := 16#B1AA;
   END_VAR
BEGIN
END_DATA_BLOCK

ORGANIZATION_BLOCK "Main"   // OB1, LAD, ProgramCycle
TITLE = "Main Program Sweep (Cycle)"
{ S7_Optimized_Access := 'TRUE' }
VERSION : 0.1
// stored: AutoNumber true, IsIECCheckEnabled false, SetENOAutomatically false
   VAR_INPUT
      Initial_Call : Bool;   // Initial call of this OB
      Remanence : Bool;   // =True, if remanent data are available
   END_VAR
   VAR_TEMP   // added for the SCL form of the ladder/FBD networks
      _w1 : Bool;
      _w2 : Bool;
      _w3 : Bool;
      _w4 : Bool;
      _w5 : Bool;
   END_VAR
BEGIN

REGION Network 1: Communication
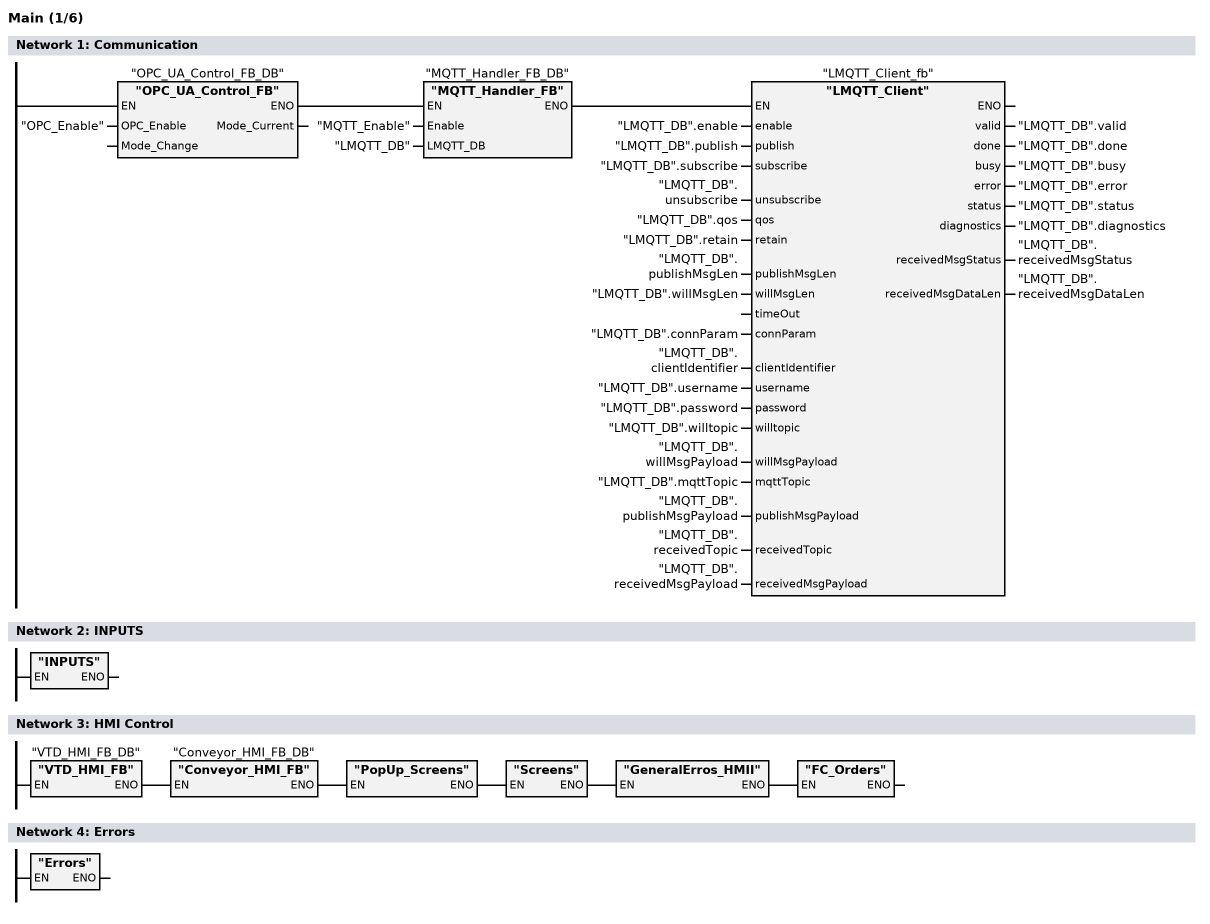
   RUNG wire#powerrail
      "OPC_UA_Control_FB_DB"(OPC_Enable := "OPC_Enable", Mode_Change :=, Mode_Current =>)
      "MQTT_Handler_FB_DB"(Enable := "MQTT_Enable", LMQTT_DB := "LMQTT_DB")
      "LMQTT_Client_fb"(enable := "LMQTT_DB".enable, publish := "LMQTT_DB".publish, subscribe := "LMQTT_DB".subscribe, unsubscribe := "LMQTT_DB".unsubscribe, qos := "LMQTT_DB".qos, retain := "LMQTT_DB".retain, publishMsgLen := "LMQTT_DB".publishMsgLen, willMsgLen := "LMQTT_DB".willMsgLen, timeOut :=, connParam := "LMQTT_DB".connParam, clientIdentifier := "LMQTT_DB".clientIdentifier, username := "LMQTT_DB".username, password := "LMQTT_DB".password, willtopic := "LMQTT_DB".willtopic, willMsgPayload := "LMQTT_DB".willMsgPayload, mqttTopic := "LMQTT_DB".mqttTopic, publishMsgPayload := "LMQTT_DB".publishMsgPayload, receivedTopic := "LMQTT_DB".receivedTopic, receivedMsgPayload := "LMQTT_DB".receivedMsgPayload, valid => "LMQTT_DB".valid, done => "LMQTT_DB".done, busy => "LMQTT_DB".busy, error => "LMQTT_DB".error, status => "LMQTT_DB".status, diagnostics => "LMQTT_DB".diagnostics, receivedMsgStatus => "LMQTT_DB".receivedMsgStatus, receivedMsgDataLen => "LMQTT_DB".receivedMsgDataLen)
   END_RUNG
   // the same network as SCL:
   "OPC_UA_Control_FB_DB"(OPC_Enable := "OPC_Enable", ENO => #_w1);   // "OPC_UA_Control_FB"
   "MQTT_Handler_FB_DB"(EN := #_w1, Enable := "MQTT_Enable", LMQTT_DB := "LMQTT_DB", ENO => #_w2);   // "MQTT_Handler_FB"
   IF #_w2 THEN
       "LMQTT_Client_fb"(enable := "LMQTT_DB".enable,   // "LMQTT_Client"
                         publish := "LMQTT_DB".publish,
                         subscribe := "LMQTT_DB".subscribe,
                         unsubscribe := "LMQTT_DB".unsubscribe,
                         qos := "LMQTT_DB".qos,
                         retain := "LMQTT_DB".retain,
                         publishMsgLen := "LMQTT_DB".publishMsgLen,
                         willMsgLen := "LMQTT_DB".willMsgLen,
                         connParam := "LMQTT_DB".connParam,
                         clientIdentifier := "LMQTT_DB".clientIdentifier,
                         username := "LMQTT_DB".username,
                         password := "LMQTT_DB".password,
                         willtopic := "LMQTT_DB".willtopic,
                         willMsgPayload := "LMQTT_DB".willMsgPayload,
                         mqttTopic := "LMQTT_DB".mqttTopic,
                         publishMsgPayload := "LMQTT_DB".publishMsgPayload,
                         receivedTopic := "LMQTT_DB".receivedTopic,
                         receivedMsgPayload := "LMQTT_DB".receivedMsgPayload,
                         valid => "LMQTT_DB".valid,
                         done => "LMQTT_DB".done,
                         busy => "LMQTT_DB".busy,
                         error => "LMQTT_DB".error,
                         status => "LMQTT_DB".status,
                         diagnostics => "LMQTT_DB".diagnostics,
                         receivedMsgStatus => "LMQTT_DB".receivedMsgStatus,
                         receivedMsgDataLen => "LMQTT_DB".receivedMsgDataLen);
   END_IF;
END_REGION

REGION Network 2: INPUTS
   RUNG wire#powerrail
      "INPUTS"()
   END_RUNG
   // the same network as SCL:
   "INPUTS"();
END_REGION

REGION Network 3: HMI Control
   RUNG wire#powerrail
      "VTD_HMI_FB_DB"()
      "Conveyor_HMI_FB_DB"()
      "PopUp_Screens"()
      "Screens"()
      "GeneralErros_HMII"()
      "FC_Orders"()
   END_RUNG
   // the same network as SCL:
   "VTD_HMI_FB_DB"(ENO => #_w1);   // "VTD_HMI_FB"
   "Conveyor_HMI_FB_DB"(EN := #_w1, ENO => #_w2);   // "Conveyor_HMI_FB"
   "PopUp_Screens"(EN := #_w2, ENO => #_w3);
   "Screens"(EN := #_w3, ENO => #_w4);
   "GeneralErros_HMII"(EN := #_w4, ENO => #_w5);
   IF #_w5 THEN "FC_Orders"(); END_IF;
END_REGION

REGION Network 4: Errors
   RUNG wire#powerrail
      "Errors"()
   END_RUNG
   // the same network as SCL:
   "Errors"();
END_REGION

REGION Network 5: Carousel Conveyors
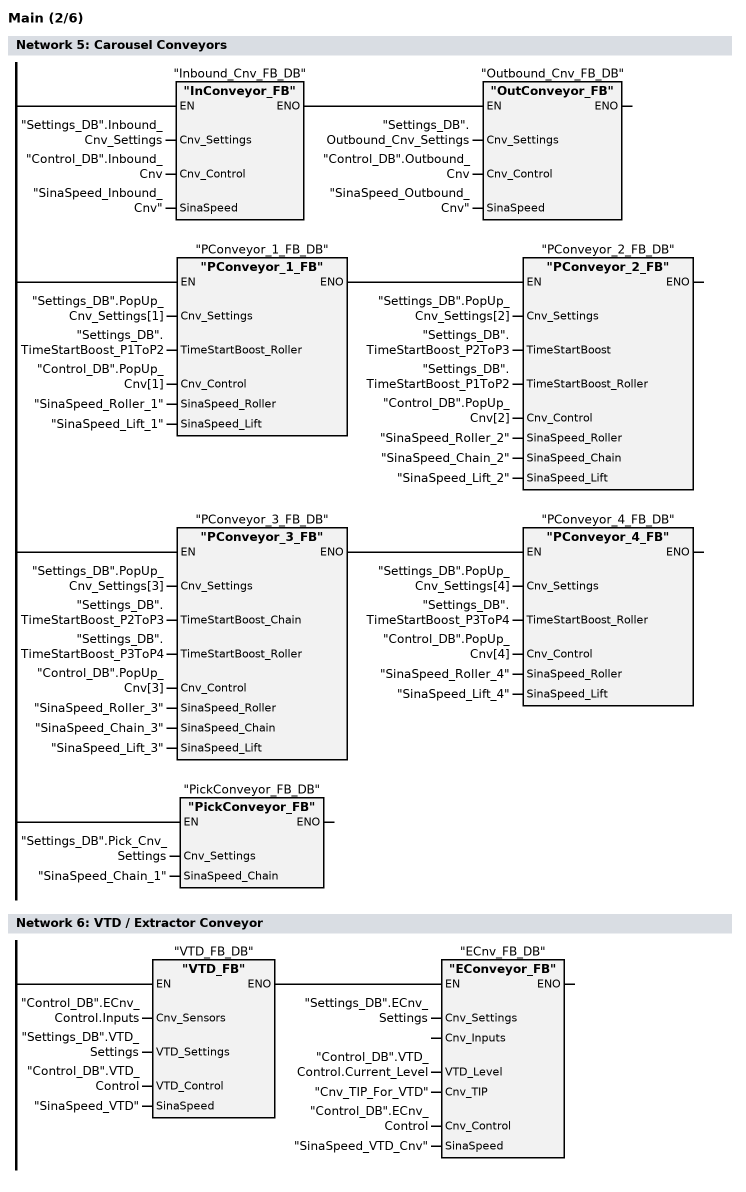
   RUNG wire#powerrail
      "Inbound_Cnv_FB_DB"(Cnv_Settings := "Settings_DB".Inbound_Cnv_Settings, Cnv_Control := "Control_DB".Inbound_Cnv, SinaSpeed := "SinaSpeed_Inbound_Cnv")
      "Outbound_Cnv_FB_DB"(Cnv_Settings := "Settings_DB".Outbound_Cnv_Settings, Cnv_Control := "Control_DB".Outbound_Cnv, SinaSpeed := "SinaSpeed_Outbound_Cnv")
   END_RUNG
   RUNG wire#powerrail
      "PConveyor_1_FB_DB"(Cnv_Settings := "Settings_DB".PopUp_Cnv_Settings[1], TimeStartBoost_Roller := "Settings_DB".TimeStartBoost_P1ToP2, Cnv_Control := "Control_DB".PopUp_Cnv[1], SinaSpeed_Roller := "SinaSpeed_Roller_1", SinaSpeed_Lift := "SinaSpeed_Lift_1")
      "PConveyor_2_FB_DB"(Cnv_Settings := "Settings_DB".PopUp_Cnv_Settings[2], TimeStartBoost := "Settings_DB".TimeStartBoost_P2ToP3, TimeStartBoost_Roller := "Settings_DB".TimeStartBoost_P1ToP2, Cnv_Control := "Control_DB".PopUp_Cnv[2], SinaSpeed_Roller := "SinaSpeed_Roller_2", SinaSpeed_Chain := "SinaSpeed_Chain_2", SinaSpeed_Lift := "SinaSpeed_Lift_2")
   END_RUNG
   RUNG wire#powerrail
      "PConveyor_3_FB_DB"(Cnv_Settings := "Settings_DB".PopUp_Cnv_Settings[3], TimeStartBoost_Chain := "Settings_DB".TimeStartBoost_P2ToP3, TimeStartBoost_Roller := "Settings_DB".TimeStartBoost_P3ToP4, Cnv_Control := "Control_DB".PopUp_Cnv[3], SinaSpeed_Roller := "SinaSpeed_Roller_3", SinaSpeed_Chain := "SinaSpeed_Chain_3", SinaSpeed_Lift := "SinaSpeed_Lift_3")
      "PConveyor_4_FB_DB"(Cnv_Settings := "Settings_DB".PopUp_Cnv_Settings[4], TimeStartBoost_Roller := "Settings_DB".TimeStartBoost_P3ToP4, Cnv_Control := "Control_DB".PopUp_Cnv[4], SinaSpeed_Roller := "SinaSpeed_Roller_4", SinaSpeed_Lift := "SinaSpeed_Lift_4")
   END_RUNG
   RUNG wire#powerrail
      "PickConveyor_FB_DB"(Cnv_Settings := "Settings_DB".Pick_Cnv_Settings, SinaSpeed_Chain := "SinaSpeed_Chain_1")
   END_RUNG
   // the same network as SCL:
   "Inbound_Cnv_FB_DB"(Cnv_Settings := "Settings_DB".Inbound_Cnv_Settings,   // "InConveyor_FB"
                       Cnv_Control := "Control_DB".Inbound_Cnv,
                       SinaSpeed := "SinaSpeed_Inbound_Cnv",
                       ENO => #_w1);
   IF #_w1 THEN
       "Outbound_Cnv_FB_DB"(Cnv_Settings := "Settings_DB".Outbound_Cnv_Settings,   // "OutConveyor_FB"
                            Cnv_Control := "Control_DB".Outbound_Cnv,
                            SinaSpeed := "SinaSpeed_Outbound_Cnv");
   END_IF;
   "PConveyor_1_FB_DB"(Cnv_Settings := "Settings_DB".PopUp_Cnv_Settings[1],   // "PConveyor_1_FB"
                       TimeStartBoost_Roller := "Settings_DB".TimeStartBoost_P1ToP2,
                       Cnv_Control := "Control_DB".PopUp_Cnv[1],
                       SinaSpeed_Roller := "SinaSpeed_Roller_1",
                       SinaSpeed_Lift := "SinaSpeed_Lift_1",
                       ENO => #_w2);
   IF #_w2 THEN
       "PConveyor_2_FB_DB"(Cnv_Settings := "Settings_DB".PopUp_Cnv_Settings[2],   // "PConveyor_2_FB"
                           TimeStartBoost := "Settings_DB".TimeStartBoost_P2ToP3,
                           TimeStartBoost_Roller := "Settings_DB".TimeStartBoost_P1ToP2,
                           Cnv_Control := "Control_DB".PopUp_Cnv[2],
                           SinaSpeed_Roller := "SinaSpeed_Roller_2",
                           SinaSpeed_Chain := "SinaSpeed_Chain_2",
                           SinaSpeed_Lift := "SinaSpeed_Lift_2");
   END_IF;
   "PConveyor_3_FB_DB"(Cnv_Settings := "Settings_DB".PopUp_Cnv_Settings[3],   // "PConveyor_3_FB"
                       TimeStartBoost_Chain := "Settings_DB".TimeStartBoost_P2ToP3,
                       TimeStartBoost_Roller := "Settings_DB".TimeStartBoost_P3ToP4,
                       Cnv_Control := "Control_DB".PopUp_Cnv[3],
                       SinaSpeed_Roller := "SinaSpeed_Roller_3",
                       SinaSpeed_Chain := "SinaSpeed_Chain_3",
                       SinaSpeed_Lift := "SinaSpeed_Lift_3",
                       ENO => #_w3);
   IF #_w3 THEN
       "PConveyor_4_FB_DB"(Cnv_Settings := "Settings_DB".PopUp_Cnv_Settings[4],   // "PConveyor_4_FB"
                           TimeStartBoost_Roller := "Settings_DB".TimeStartBoost_P3ToP4,
                           Cnv_Control := "Control_DB".PopUp_Cnv[4],
                           SinaSpeed_Roller := "SinaSpeed_Roller_4",
                           SinaSpeed_Lift := "SinaSpeed_Lift_4");
   END_IF;
   "PickConveyor_FB_DB"(Cnv_Settings := "Settings_DB".Pick_Cnv_Settings, SinaSpeed_Chain := "SinaSpeed_Chain_1");   // "PickConveyor_FB"
END_REGION

REGION Network 6: VTD / Extractor Conveyor
   RUNG wire#powerrail
      "VTD_FB_DB"(Cnv_Sensors := "Control_DB".ECnv_Control.Inputs, VTD_Settings := "Settings_DB".VTD_Settings, VTD_Control := "Control_DB".VTD_Control, SinaSpeed := "SinaSpeed_VTD")
      "ECnv_FB_DB"(Cnv_Settings := "Settings_DB".ECnv_Settings, Cnv_Inputs :=, VTD_Level := "Control_DB".VTD_Control.Current_Level, Cnv_TIP := "Cnv_TIP_For_VTD", Cnv_Control := "Control_DB".ECnv_Control, SinaSpeed := "SinaSpeed_VTD_Cnv")
   END_RUNG
   // the same network as SCL:
   "VTD_FB_DB"(Cnv_Sensors := "Control_DB".ECnv_Control.Inputs,   // "VTD_FB"
               VTD_Settings := "Settings_DB".VTD_Settings,
               VTD_Control := "Control_DB".VTD_Control,
               SinaSpeed := "SinaSpeed_VTD",
               ENO => #_w1);
   IF #_w1 THEN
       "ECnv_FB_DB"(Cnv_Settings := "Settings_DB".ECnv_Settings,   // "EConveyor_FB"
                    VTD_Level := "Control_DB".VTD_Control.Current_Level,
                    Cnv_TIP := "Cnv_TIP_For_VTD",
                    Cnv_Control := "Control_DB".ECnv_Control,
                    SinaSpeed := "SinaSpeed_VTD_Cnv");
   END_IF;
END_REGION

REGION Network 7: Level Conveyors
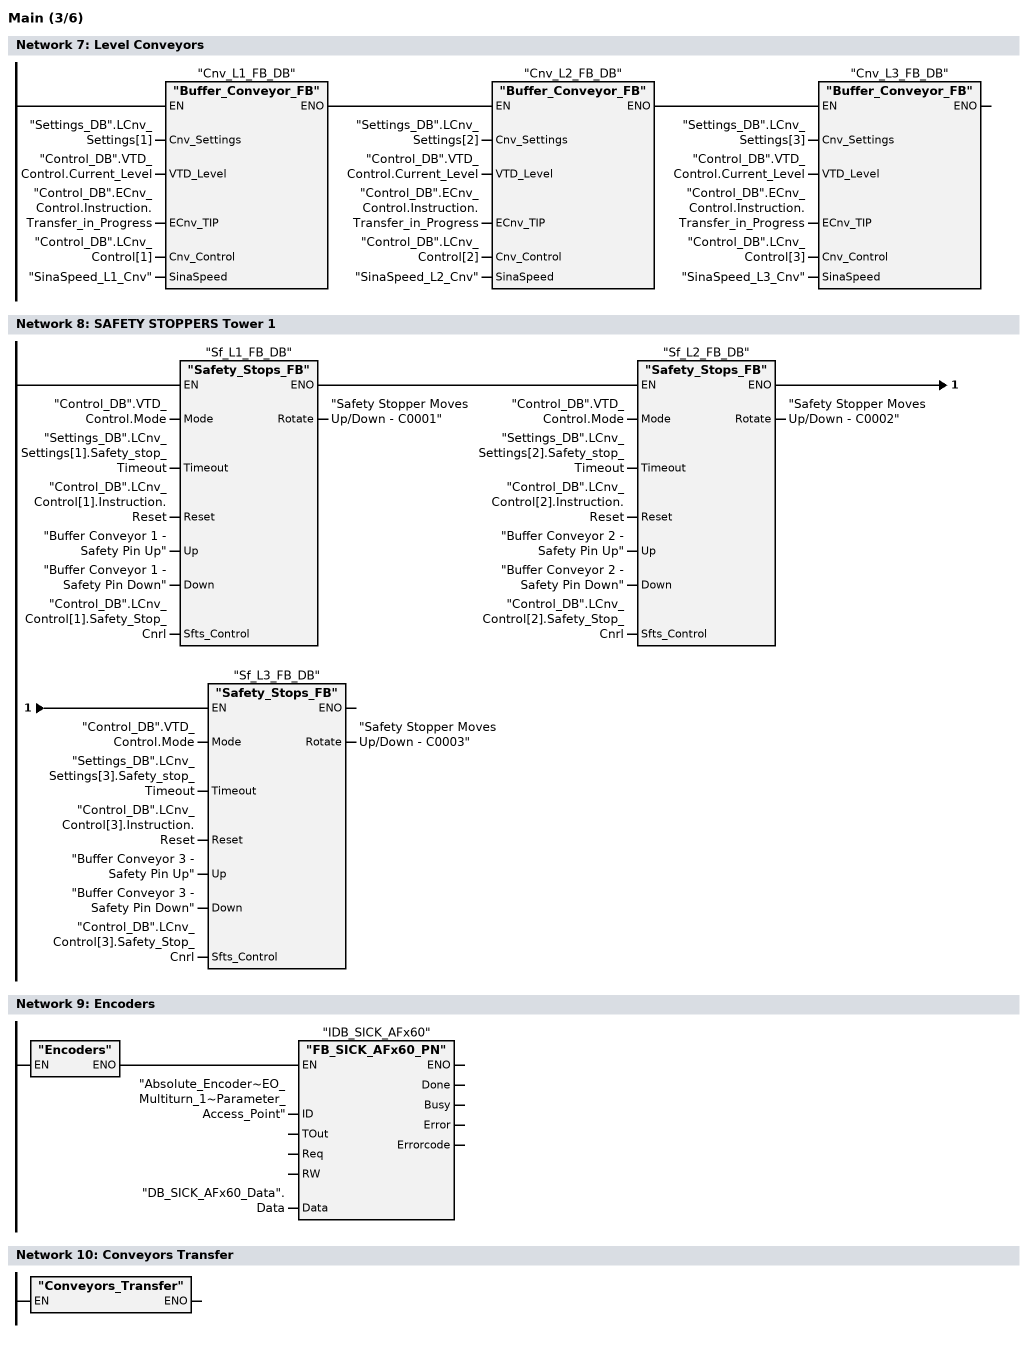
   RUNG wire#powerrail
      "Cnv_L1_FB_DB"(Cnv_Settings := "Settings_DB".LCnv_Settings[1], VTD_Level := "Control_DB".VTD_Control.Current_Level, ECnv_TIP := "Control_DB".ECnv_Control.Instruction.Transfer_in_Progress, Cnv_Control := "Control_DB".LCnv_Control[1], SinaSpeed := "SinaSpeed_L1_Cnv")
      "Cnv_L2_FB_DB"(Cnv_Settings := "Settings_DB".LCnv_Settings[2], VTD_Level := "Control_DB".VTD_Control.Current_Level, ECnv_TIP := "Control_DB".ECnv_Control.Instruction.Transfer_in_Progress, Cnv_Control := "Control_DB".LCnv_Control[2], SinaSpeed := "SinaSpeed_L2_Cnv")
      "Cnv_L3_FB_DB"(Cnv_Settings := "Settings_DB".LCnv_Settings[3], VTD_Level := "Control_DB".VTD_Control.Current_Level, ECnv_TIP := "Control_DB".ECnv_Control.Instruction.Transfer_in_Progress, Cnv_Control := "Control_DB".LCnv_Control[3], SinaSpeed := "SinaSpeed_L3_Cnv")
   END_RUNG
   // the same network as SCL:
   "Cnv_L1_FB_DB"(Cnv_Settings := "Settings_DB".LCnv_Settings[1],   // "Buffer_Conveyor_FB"
                  VTD_Level := "Control_DB".VTD_Control.Current_Level,
                  ECnv_TIP := "Control_DB".ECnv_Control.Instruction.Transfer_in_Progress,
                  Cnv_Control := "Control_DB".LCnv_Control[1],
                  SinaSpeed := "SinaSpeed_L1_Cnv",
                  ENO => #_w1);
   "Cnv_L2_FB_DB"(EN := #_w1,   // "Buffer_Conveyor_FB"
                  Cnv_Settings := "Settings_DB".LCnv_Settings[2],
                  VTD_Level := "Control_DB".VTD_Control.Current_Level,
                  ECnv_TIP := "Control_DB".ECnv_Control.Instruction.Transfer_in_Progress,
                  Cnv_Control := "Control_DB".LCnv_Control[2],
                  SinaSpeed := "SinaSpeed_L2_Cnv",
                  ENO => #_w2);
   IF #_w2 THEN
       "Cnv_L3_FB_DB"(Cnv_Settings := "Settings_DB".LCnv_Settings[3],   // "Buffer_Conveyor_FB"
                      VTD_Level := "Control_DB".VTD_Control.Current_Level,
                      ECnv_TIP := "Control_DB".ECnv_Control.Instruction.Transfer_in_Progress,
                      Cnv_Control := "Control_DB".LCnv_Control[3],
                      SinaSpeed := "SinaSpeed_L3_Cnv");
   END_IF;
END_REGION

REGION Network 8: SAFETY STOPPERS Tower 1
   RUNG wire#powerrail
      "Sf_L1_FB_DB"(Mode := "Control_DB".VTD_Control.Mode, Timeout := "Settings_DB".LCnv_Settings[1].Safety_stop_Timeout, Reset := "Control_DB".LCnv_Control[1].Instruction.Reset, Up := "Buffer Conveyor 1 - Safety Pin Up", Down := "Buffer Conveyor 1 - Safety Pin Down", Sfts_Control := "Control_DB".LCnv_Control[1].Safety_Stop_Cnrl, Rotate => "Safety Stopper Moves Up/Down - C0001")
      "Sf_L2_FB_DB"(Mode := "Control_DB".VTD_Control.Mode, Timeout := "Settings_DB".LCnv_Settings[2].Safety_stop_Timeout, Reset := "Control_DB".LCnv_Control[2].Instruction.Reset, Up := "Buffer Conveyor 2 - Safety Pin Up", Down := "Buffer Conveyor 2 - Safety Pin Down", Sfts_Control := "Control_DB".LCnv_Control[2].Safety_Stop_Cnrl, Rotate => "Safety Stopper Moves Up/Down - C0002")
      "Sf_L3_FB_DB"(Mode := "Control_DB".VTD_Control.Mode, Timeout := "Settings_DB".LCnv_Settings[3].Safety_stop_Timeout, Reset := "Control_DB".LCnv_Control[3].Instruction.Reset, Up := "Buffer Conveyor 3 - Safety Pin Up", Down := "Buffer Conveyor 3 - Safety Pin Down", Sfts_Control := "Control_DB".LCnv_Control[3].Safety_Stop_Cnrl, Rotate => "Safety Stopper Moves Up/Down - C0003")
   END_RUNG
   // the same network as SCL:
   "Sf_L1_FB_DB"(Mode := "Control_DB".VTD_Control.Mode,   // "Safety_Stops_FB"
                 Timeout := "Settings_DB".LCnv_Settings[1].Safety_stop_Timeout,
                 Reset := "Control_DB".LCnv_Control[1].Instruction.Reset,
                 Up := "Buffer Conveyor 1 - Safety Pin Up",
                 Down := "Buffer Conveyor 1 - Safety Pin Down",
                 Sfts_Control := "Control_DB".LCnv_Control[1].Safety_Stop_Cnrl,
                 Rotate => "Safety Stopper Moves Up/Down - C0001",
                 ENO => #_w1);
   "Sf_L2_FB_DB"(EN := #_w1,   // "Safety_Stops_FB"
                 Mode := "Control_DB".VTD_Control.Mode,
                 Timeout := "Settings_DB".LCnv_Settings[2].Safety_stop_Timeout,
                 Reset := "Control_DB".LCnv_Control[2].Instruction.Reset,
                 Up := "Buffer Conveyor 2 - Safety Pin Up",
                 Down := "Buffer Conveyor 2 - Safety Pin Down",
                 Sfts_Control := "Control_DB".LCnv_Control[2].Safety_Stop_Cnrl,
                 Rotate => "Safety Stopper Moves Up/Down - C0002",
                 ENO => #_w2);
   IF #_w2 THEN
       "Sf_L3_FB_DB"(Mode := "Control_DB".VTD_Control.Mode,   // "Safety_Stops_FB"
                     Timeout := "Settings_DB".LCnv_Settings[3].Safety_stop_Timeout,
                     Reset := "Control_DB".LCnv_Control[3].Instruction.Reset,
                     Up := "Buffer Conveyor 3 - Safety Pin Up",
                     Down := "Buffer Conveyor 3 - Safety Pin Down",
                     Sfts_Control := "Control_DB".LCnv_Control[3].Safety_Stop_Cnrl,
                     Rotate => "Safety Stopper Moves Up/Down - C0003");
   END_IF;
END_REGION

REGION Network 9: Encoders
   RUNG wire#powerrail
      "Encoders"()
      "IDB_SICK_AFx60"(ID := "Absolute_Encoder~EO_Multiturn_1~Parameter_Access_Point", TOut :=, Req :=, RW :=, Data := "DB_SICK_AFx60_Data".Data, Done =>, Busy =>, Error =>, Errorcode =>)
   END_RUNG
   // the same network as SCL:
   "Encoders"(ENO => #_w1);
   IF #_w1 THEN
       "IDB_SICK_AFx60"(ID := "Absolute_Encoder~EO_Multiturn_1~Parameter_Access_Point",   // "FB_SICK_AFx60_PN"
                        Data := "DB_SICK_AFx60_Data".Data);
   END_IF;
END_REGION

REGION Network 10: Conveyors Transfer
   RUNG wire#powerrail
      "Conveyors_Transfer"()
   END_RUNG
   // the same network as SCL:
   "Conveyors_Transfer"();
END_REGION

REGION Network 11: Lightbar
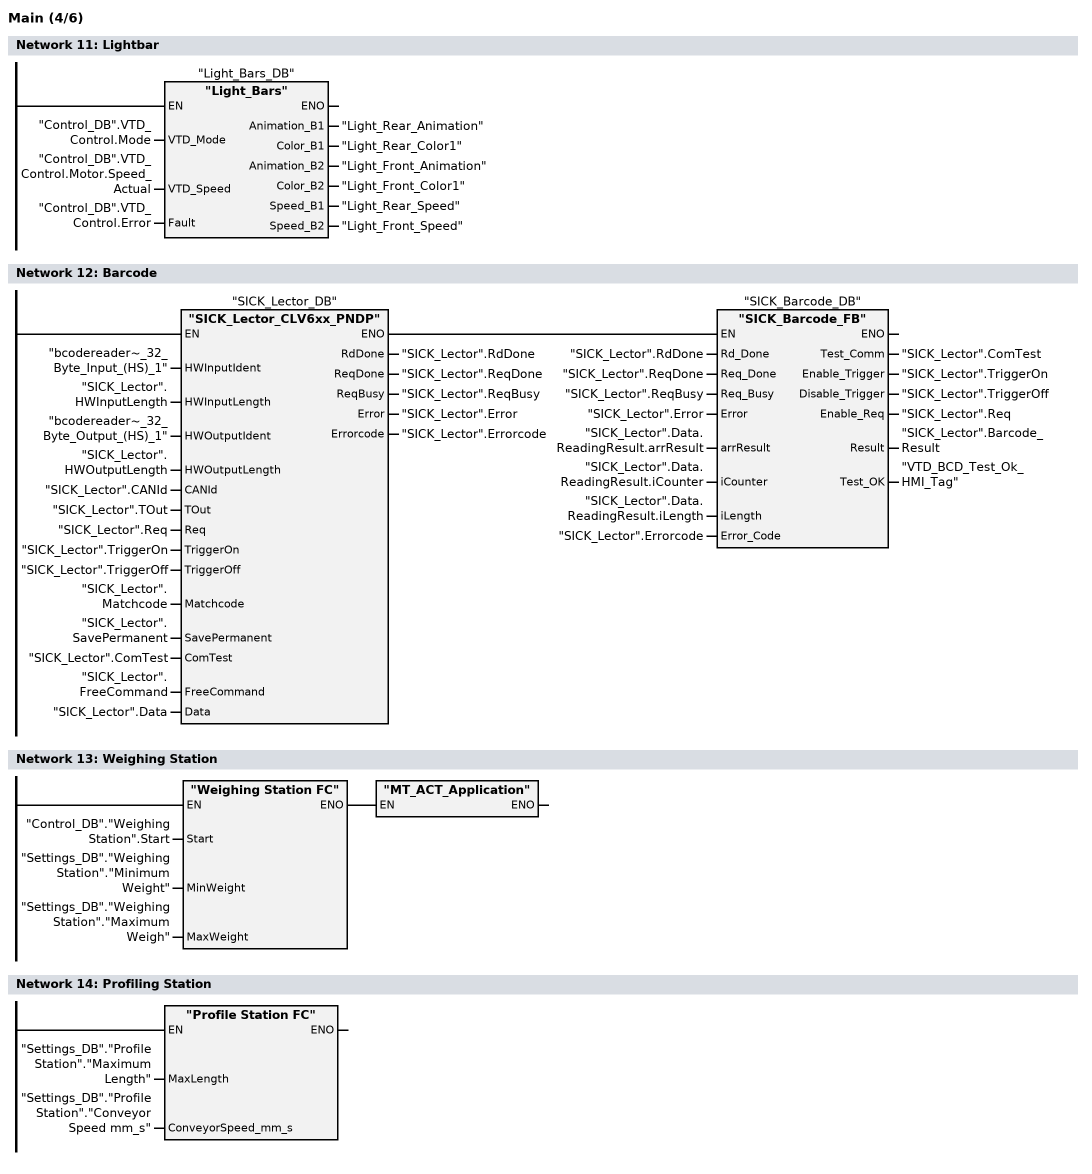
   RUNG wire#powerrail
      "Light_Bars_DB"(VTD_Mode := "Control_DB".VTD_Control.Mode, VTD_Speed := "Control_DB".VTD_Control.Motor.Speed_Actual, Fault := "Control_DB".VTD_Control.Error, Animation_B1 => "Light_Rear_Animation", Color_B1 => "Light_Rear_Color1", Animation_B2 => "Light_Front_Animation", Color_B2 => "Light_Front_Color1", Speed_B1 => "Light_Rear_Speed", Speed_B2 => "Light_Front_Speed")
   END_RUNG
   // the same network as SCL:
   "Light_Bars_DB"(VTD_Mode := "Control_DB".VTD_Control.Mode,   // "Light_Bars"
                   VTD_Speed := "Control_DB".VTD_Control.Motor.Speed_Actual,
                   Fault := "Control_DB".VTD_Control.Error,
                   Animation_B1 => "Light_Rear_Animation",
                   Color_B1 => "Light_Rear_Color1",
                   Animation_B2 => "Light_Front_Animation",
                   Color_B2 => "Light_Front_Color1",
                   Speed_B1 => "Light_Rear_Speed",
                   Speed_B2 => "Light_Front_Speed");
END_REGION

REGION Network 12: Barcode
   RUNG wire#powerrail
      "SICK_Lector_DB"(HWInputIdent := "bcodereader~_32_Byte_Input_(HS)_1", HWInputLength := "SICK_Lector".HWInputLength, HWOutputIdent := "bcodereader~_32_Byte_Output_(HS)_1", HWOutputLength := "SICK_Lector".HWOutputLength, CANId := "SICK_Lector".CANId, TOut := "SICK_Lector".TOut, Req := "SICK_Lector".Req, TriggerOn := "SICK_Lector".TriggerOn, TriggerOff := "SICK_Lector".TriggerOff, Matchcode := "SICK_Lector".Matchcode, SavePermanent := "SICK_Lector".SavePermanent, ComTest := "SICK_Lector".ComTest, FreeCommand := "SICK_Lector".FreeCommand, Data := "SICK_Lector".Data, RdDone => "SICK_Lector".RdDone, ReqDone => "SICK_Lector".ReqDone, ReqBusy => "SICK_Lector".ReqBusy, Error => "SICK_Lector".Error, Errorcode => "SICK_Lector".Errorcode)
      "SICK_Barcode_DB"(Rd_Done := "SICK_Lector".RdDone, Req_Done := "SICK_Lector".ReqDone, Req_Busy := "SICK_Lector".ReqBusy, Error := "SICK_Lector".Error, arrResult := "SICK_Lector".Data.ReadingResult.arrResult, iCounter := "SICK_Lector".Data.ReadingResult.iCounter, iLength := "SICK_Lector".Data.ReadingResult.iLength, Error_Code := "SICK_Lector".Errorcode, Test_Comm => "SICK_Lector".ComTest, Enable_Trigger => "SICK_Lector".TriggerOn, Disable_Trigger => "SICK_Lector".TriggerOff, Enable_Req => "SICK_Lector".Req, Result => "SICK_Lector".Barcode_Result, Test_OK => "VTD_BCD_Test_Ok_HMI_Tag")
   END_RUNG
   // the same network as SCL:
   "SICK_Lector_DB"(HWInputIdent := "bcodereader~_32_Byte_Input_(HS)_1",   // "SICK_Lector_CLV6xx_PNDP"
                    HWInputLength := "SICK_Lector".HWInputLength,
                    HWOutputIdent := "bcodereader~_32_Byte_Output_(HS)_1",
                    HWOutputLength := "SICK_Lector".HWOutputLength,
                    CANId := "SICK_Lector".CANId,
                    TOut := "SICK_Lector".TOut,
                    Req := "SICK_Lector".Req,
                    TriggerOn := "SICK_Lector".TriggerOn,
                    TriggerOff := "SICK_Lector".TriggerOff,
                    Matchcode := "SICK_Lector".Matchcode,
                    SavePermanent := "SICK_Lector".SavePermanent,
                    ComTest := "SICK_Lector".ComTest,
                    FreeCommand := "SICK_Lector".FreeCommand,
                    Data := "SICK_Lector".Data,
                    RdDone => "SICK_Lector".RdDone,
                    ReqDone => "SICK_Lector".ReqDone,
                    ReqBusy => "SICK_Lector".ReqBusy,
                    Error => "SICK_Lector".Error,
                    Errorcode => "SICK_Lector".Errorcode,
                    ENO => #_w1);
   IF #_w1 THEN
       "SICK_Barcode_DB"(Rd_Done := "SICK_Lector".RdDone,   // "SICK_Barcode_FB"
                         Req_Done := "SICK_Lector".ReqDone,
                         Req_Busy := "SICK_Lector".ReqBusy,
                         Error := "SICK_Lector".Error,
                         arrResult := "SICK_Lector".Data.ReadingResult.arrResult,
                         iCounter := "SICK_Lector".Data.ReadingResult.iCounter,
                         iLength := "SICK_Lector".Data.ReadingResult.iLength,
                         Error_Code := "SICK_Lector".Errorcode,
                         Test_Comm => "SICK_Lector".ComTest,
                         Enable_Trigger => "SICK_Lector".TriggerOn,
                         Disable_Trigger => "SICK_Lector".TriggerOff,
                         Enable_Req => "SICK_Lector".Req,
                         Result => "SICK_Lector".Barcode_Result,
                         Test_OK => "VTD_BCD_Test_Ok_HMI_Tag");
   END_IF;
END_REGION

REGION Network 13: Weighing Station
   RUNG wire#powerrail
      "Weighing Station FC"(Start := "Control_DB"."Weighing Station".Start, MinWeight := "Settings_DB"."Weighing Station"."Minimum Weight", MaxWeight := "Settings_DB"."Weighing Station"."Maximum Weigh")
      "MT_ACT_Application"()
   END_RUNG
   // the same network as SCL:
   "Weighing Station FC"(Start := "Control_DB"."Weighing Station".Start,
                         MinWeight := "Settings_DB"."Weighing Station"."Minimum Weight",
                         MaxWeight := "Settings_DB"."Weighing Station"."Maximum Weigh",
                         ENO => #_w1);
   IF #_w1 THEN "MT_ACT_Application"(); END_IF;
END_REGION

REGION Network 14: Profiling Station
   RUNG wire#powerrail
      "Profile Station FC"(MaxLength := "Settings_DB"."Profile Station"."Maximum Length", ConveyorSpeed_mm_s := "Settings_DB"."Profile Station"."Conveyor Speed mm_s")
   END_RUNG
   // the same network as SCL:
   "Profile Station FC"(MaxLength := "Settings_DB"."Profile Station"."Maximum Length",
                        ConveyorSpeed_mm_s := "Settings_DB"."Profile Station"."Conveyor Speed mm_s");
END_REGION

REGION Network 15: Barcode Stations
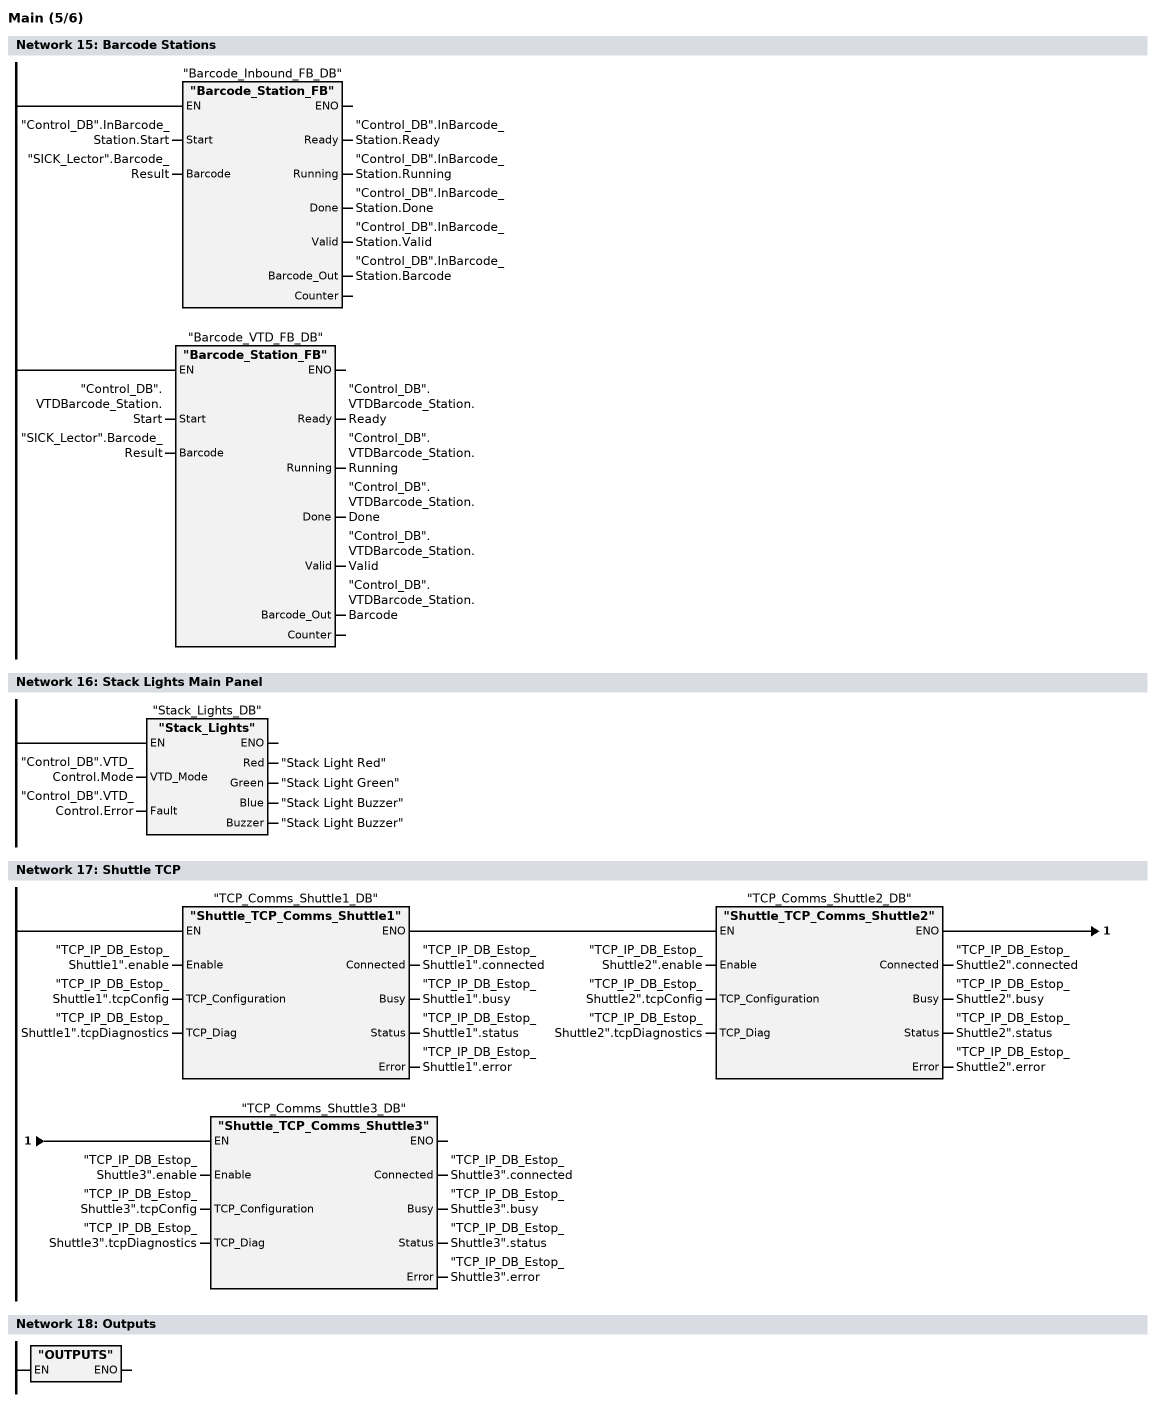
   RUNG wire#powerrail
      "Barcode_Inbound_FB_DB"(Start := "Control_DB".InBarcode_Station.Start, Barcode := "SICK_Lector".Barcode_Result, Ready => "Control_DB".InBarcode_Station.Ready, Running => "Control_DB".InBarcode_Station.Running, Done => "Control_DB".InBarcode_Station.Done, Valid => "Control_DB".InBarcode_Station.Valid, Barcode_Out => "Control_DB".InBarcode_Station.Barcode, "Counter" =>)
   END_RUNG
   RUNG wire#powerrail
      "Barcode_VTD_FB_DB"(Start := "Control_DB".VTDBarcode_Station.Start, Barcode := "SICK_Lector".Barcode_Result, Ready => "Control_DB".VTDBarcode_Station.Ready, Running => "Control_DB".VTDBarcode_Station.Running, Done => "Control_DB".VTDBarcode_Station.Done, Valid => "Control_DB".VTDBarcode_Station.Valid, Barcode_Out => "Control_DB".VTDBarcode_Station.Barcode, "Counter" =>)
   END_RUNG
   // the same network as SCL:
   "Barcode_Inbound_FB_DB"(Start := "Control_DB".InBarcode_Station.Start,   // "Barcode_Station_FB"
                           Barcode := "SICK_Lector".Barcode_Result,
                           Ready => "Control_DB".InBarcode_Station.Ready,
                           Running => "Control_DB".InBarcode_Station.Running,
                           Done => "Control_DB".InBarcode_Station.Done,
                           Valid => "Control_DB".InBarcode_Station.Valid,
                           Barcode_Out => "Control_DB".InBarcode_Station.Barcode);
   "Barcode_VTD_FB_DB"(Start := "Control_DB".VTDBarcode_Station.Start,   // "Barcode_Station_FB"
                       Barcode := "SICK_Lector".Barcode_Result,
                       Ready => "Control_DB".VTDBarcode_Station.Ready,
                       Running => "Control_DB".VTDBarcode_Station.Running,
                       Done => "Control_DB".VTDBarcode_Station.Done,
                       Valid => "Control_DB".VTDBarcode_Station.Valid,
                       Barcode_Out => "Control_DB".VTDBarcode_Station.Barcode);
END_REGION

REGION Network 16: Stack Lights Main Panel
   RUNG wire#powerrail
      "Stack_Lights_DB"(VTD_Mode := "Control_DB".VTD_Control.Mode, Fault := "Control_DB".VTD_Control.Error, Red => "Stack Light Red", Green => "Stack Light Green", Blue => "Stack Light Buzzer", Buzzer => "Stack Light Buzzer")
   END_RUNG
   // the same network as SCL:
   "Stack_Lights_DB"(VTD_Mode := "Control_DB".VTD_Control.Mode,   // "Stack_Lights"
                     Fault := "Control_DB".VTD_Control.Error,
                     Red => "Stack Light Red",
                     Green => "Stack Light Green",
                     Blue => "Stack Light Buzzer",
                     Buzzer => "Stack Light Buzzer");
END_REGION

REGION Network 17: Shuttle TCP
   RUNG wire#powerrail
      "TCP_Comms_Shuttle1_DB"(Enable := "TCP_IP_DB_Estop_Shuttle1".enable, TCP_Configuration := "TCP_IP_DB_Estop_Shuttle1".tcpConfig, TCP_Diag := "TCP_IP_DB_Estop_Shuttle1".tcpDiagnostics, Connected => "TCP_IP_DB_Estop_Shuttle1".connected, Busy => "TCP_IP_DB_Estop_Shuttle1".busy, Status => "TCP_IP_DB_Estop_Shuttle1".status, Error => "TCP_IP_DB_Estop_Shuttle1".error)
      "TCP_Comms_Shuttle2_DB"(Enable := "TCP_IP_DB_Estop_Shuttle2".enable, TCP_Configuration := "TCP_IP_DB_Estop_Shuttle2".tcpConfig, TCP_Diag := "TCP_IP_DB_Estop_Shuttle2".tcpDiagnostics, Connected => "TCP_IP_DB_Estop_Shuttle2".connected, Busy => "TCP_IP_DB_Estop_Shuttle2".busy, Status => "TCP_IP_DB_Estop_Shuttle2".status, Error => "TCP_IP_DB_Estop_Shuttle2".error)
      "TCP_Comms_Shuttle3_DB"(Enable := "TCP_IP_DB_Estop_Shuttle3".enable, TCP_Configuration := "TCP_IP_DB_Estop_Shuttle3".tcpConfig, TCP_Diag := "TCP_IP_DB_Estop_Shuttle3".tcpDiagnostics, Connected => "TCP_IP_DB_Estop_Shuttle3".connected, Busy => "TCP_IP_DB_Estop_Shuttle3".busy, Status => "TCP_IP_DB_Estop_Shuttle3".status, Error => "TCP_IP_DB_Estop_Shuttle3".error)
   END_RUNG
   // the same network as SCL:
   "TCP_Comms_Shuttle1_DB"(Enable := "TCP_IP_DB_Estop_Shuttle1".enable,   // "Shuttle_TCP_Comms_Shuttle1"
                           TCP_Configuration := "TCP_IP_DB_Estop_Shuttle1".tcpConfig,
                           TCP_Diag := "TCP_IP_DB_Estop_Shuttle1".tcpDiagnostics,
                           Connected => "TCP_IP_DB_Estop_Shuttle1".connected,
                           Busy => "TCP_IP_DB_Estop_Shuttle1".busy,
                           Status => "TCP_IP_DB_Estop_Shuttle1".status,
                           Error => "TCP_IP_DB_Estop_Shuttle1".error,
                           ENO => #_w1);
   "TCP_Comms_Shuttle2_DB"(EN := #_w1,   // "Shuttle_TCP_Comms_Shuttle2"
                           Enable := "TCP_IP_DB_Estop_Shuttle2".enable,
                           TCP_Configuration := "TCP_IP_DB_Estop_Shuttle2".tcpConfig,
                           TCP_Diag := "TCP_IP_DB_Estop_Shuttle2".tcpDiagnostics,
                           Connected => "TCP_IP_DB_Estop_Shuttle2".connected,
                           Busy => "TCP_IP_DB_Estop_Shuttle2".busy,
                           Status => "TCP_IP_DB_Estop_Shuttle2".status,
                           Error => "TCP_IP_DB_Estop_Shuttle2".error,
                           ENO => #_w2);
   IF #_w2 THEN
       "TCP_Comms_Shuttle3_DB"(Enable := "TCP_IP_DB_Estop_Shuttle3".enable,   // "Shuttle_TCP_Comms_Shuttle3"
                               TCP_Configuration := "TCP_IP_DB_Estop_Shuttle3".tcpConfig,
                               TCP_Diag := "TCP_IP_DB_Estop_Shuttle3".tcpDiagnostics,
                               Connected => "TCP_IP_DB_Estop_Shuttle3".connected,
                               Busy => "TCP_IP_DB_Estop_Shuttle3".busy,
                               Status => "TCP_IP_DB_Estop_Shuttle3".status,
                               Error => "TCP_IP_DB_Estop_Shuttle3".error);
   END_IF;
END_REGION

REGION Network 18: Outputs
   RUNG wire#powerrail
      "OUTPUTS"()
   END_RUNG
   // the same network as SCL:
   "OUTPUTS"();
END_REGION

REGION Network 19: System Order Table - Carousel
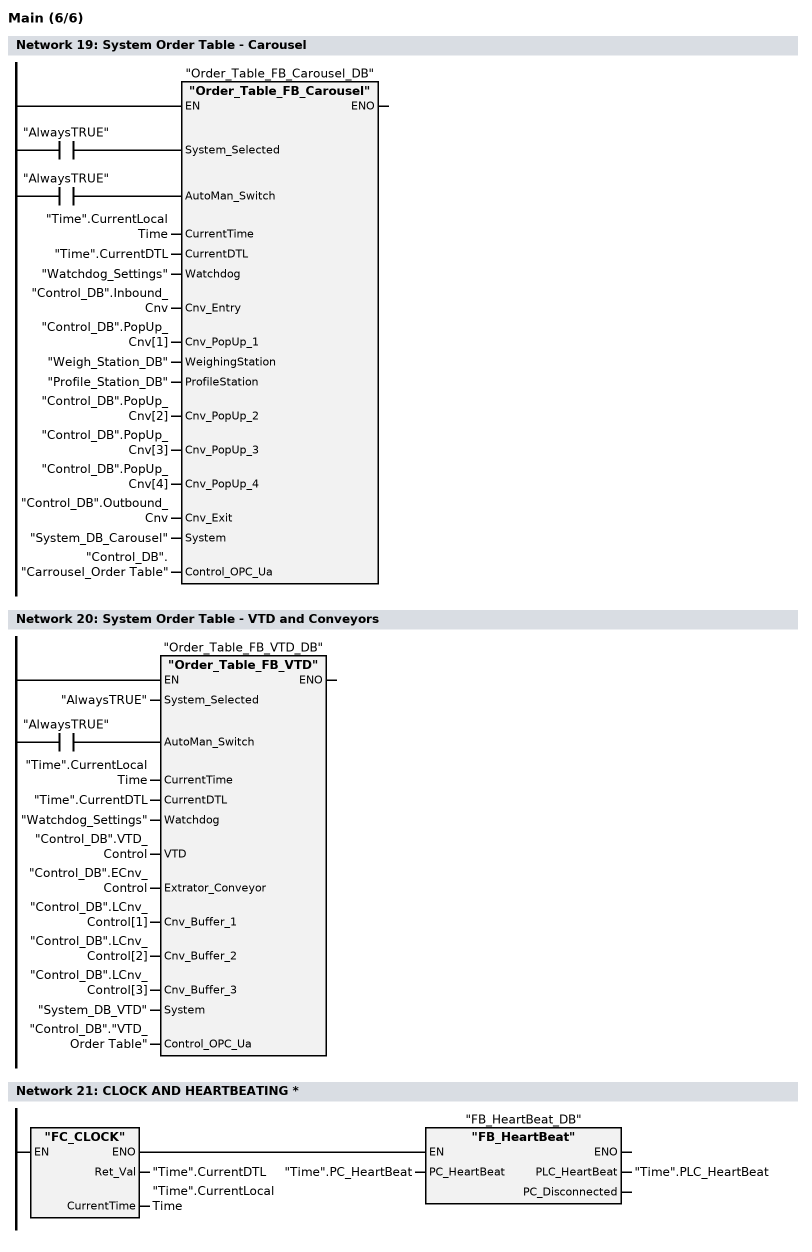
   RUNG wire#powerrail
      "Order_Table_FB_Carousel_DB"(System_Selected := wire#w1, AutoMan_Switch := wire#w2, CurrentTime := "Time".CurrentLocalTime, CurrentDTL := "Time".CurrentDTL, Watchdog := "Watchdog_Settings", Cnv_Entry := "Control_DB".Inbound_Cnv, Cnv_PopUp_1 := "Control_DB".PopUp_Cnv[1], WeighingStation := "Weigh_Station_DB", ProfileStation := "Profile_Station_DB", Cnv_PopUp_2 := "Control_DB".PopUp_Cnv[2], Cnv_PopUp_3 := "Control_DB".PopUp_Cnv[3], Cnv_PopUp_4 := "Control_DB".PopUp_Cnv[4], Cnv_Exit := "Control_DB".Outbound_Cnv, System := "System_DB_Carousel", Control_OPC_Ua := "Control_DB"."Carrousel_Order Table")
   END_RUNG
   RUNG wire#powerrail
      Contact( "AlwaysTRUE" )
   END_RUNG wire#w1
   RUNG wire#powerrail
      Contact( "AlwaysTRUE" )
   END_RUNG wire#w2
   // the same network as SCL:
   "Order_Table_FB_Carousel_DB"(System_Selected := "AlwaysTRUE",   // "Order_Table_FB_Carousel"
                           AutoMan_Switch := "AlwaysTRUE",
                           CurrentTime := "Time".CurrentLocalTime,
                           CurrentDTL := "Time".CurrentDTL,
                           Watchdog := "Watchdog_Settings",
                           Cnv_Entry := "Control_DB".Inbound_Cnv,
                           Cnv_PopUp_1 := "Control_DB".PopUp_Cnv[1],
                           WeighingStation := "Weigh_Station_DB",
                           ProfileStation := "Profile_Station_DB",
                           Cnv_PopUp_2 := "Control_DB".PopUp_Cnv[2],
                           Cnv_PopUp_3 := "Control_DB".PopUp_Cnv[3],
                           Cnv_PopUp_4 := "Control_DB".PopUp_Cnv[4],
                           Cnv_Exit := "Control_DB".Outbound_Cnv,
                           System := "System_DB_Carousel",
                           Control_OPC_Ua := "Control_DB"."Carrousel_Order Table");
END_REGION

REGION Network 20: System Order Table - VTD and Conveyors
   RUNG wire#powerrail
      "Order_Table_FB_VTD_DB"(AutoMan_Switch := wire#w1, System_Selected := "AlwaysTRUE", CurrentTime := "Time".CurrentLocalTime, CurrentDTL := "Time".CurrentDTL, Watchdog := "Watchdog_Settings", VTD := "Control_DB".VTD_Control, Extrator_Conveyor := "Control_DB".ECnv_Control, Cnv_Buffer_1 := "Control_DB".LCnv_Control[1], Cnv_Buffer_2 := "Control_DB".LCnv_Control[2], Cnv_Buffer_3 := "Control_DB".LCnv_Control[3], System := "System_DB_VTD", Control_OPC_Ua := "Control_DB"."VTD_Order Table")
   END_RUNG
   RUNG wire#powerrail
      Contact( "AlwaysTRUE" )
   END_RUNG wire#w1
   // the same network as SCL:
   "Order_Table_FB_VTD_DB"(System_Selected := "AlwaysTRUE",   // "Order_Table_FB_VTD"
                           AutoMan_Switch := "AlwaysTRUE",
                           CurrentTime := "Time".CurrentLocalTime,
                           CurrentDTL := "Time".CurrentDTL,
                           Watchdog := "Watchdog_Settings",
                           VTD := "Control_DB".VTD_Control,
                           Extrator_Conveyor := "Control_DB".ECnv_Control,
                           Cnv_Buffer_1 := "Control_DB".LCnv_Control[1],
                           Cnv_Buffer_2 := "Control_DB".LCnv_Control[2],
                           Cnv_Buffer_3 := "Control_DB".LCnv_Control[3],
                           System := "System_DB_VTD",
                           Control_OPC_Ua := "Control_DB"."VTD_Order Table");
END_REGION

REGION Network 21: CLOCK AND HEARTBEATING *
   RUNG wire#powerrail
      "FC_CLOCK"(Ret_Val => "Time".CurrentDTL, CurrentTime => "Time".CurrentLocalTime)
      "FB_HeartBeat_DB"(PC_HeartBeat := "Time".PC_HeartBeat, PLC_HeartBeat => "Time".PLC_HeartBeat, PC_Disconnected =>)
   END_RUNG
   // the same network as SCL:
   "Time".CurrentDTL := "FC_CLOCK"(CurrentTime => "Time".CurrentLocalTime, ENO => #_w1);
   IF #_w1 THEN
       "FB_HeartBeat_DB"(PC_HeartBeat := "Time".PC_HeartBeat, PLC_HeartBeat => "Time".PLC_HeartBeat);   // "FB_HeartBeat"
   END_IF;
END_REGION
END_ORGANIZATION_BLOCK

FUNCTION_BLOCK "OPC_UA_Control_FB"   // FB8, SCL
{ S7_Optimized_Access := 'TRUE' }
VERSION : 0.1
// stored: AutoNumber true, IsIECCheckEnabled false, IsRetainMemResEnabled false, MemoryReserve 100, SetENOAutomatically false, UDAEnableTagReadback false
   VAR_INPUT
      OPC_Enable : Bool;
      Mode_Change : UInt;
   END_VAR
   VAR_OUTPUT
      Mode_Current : UInt;
   END_VAR
   VAR
      Source_Location_VTD { ExternalAccessible := 'False'; ExternalVisible := 'False'; ExternalWritable := 'False'} : "ID_Decoded";
      Destination_Location_VTD { ExternalAccessible := 'False'; ExternalVisible := 'False'; ExternalWritable := 'False'} : "ID_Decoded";
      Source_Location_Carousel { ExternalAccessible := 'False'; ExternalVisible := 'False'; ExternalWritable := 'False'} : "ID_Decoded";
      Destination_Location_Carousel { ExternalAccessible := 'False'; ExternalVisible := 'False'; ExternalWritable := 'False'} : "ID_Decoded";
      State_VTD : UInt;
      State_Carrousel_Weigh : UInt;
      State_Carrousel_Main : UInt;
      State_Carrousel_PICKTP1 : UInt;
      State_Carrousel_P4TPICK : UInt;
      State_Carrousel_CTC : UInt;
      State_Carrousel_ITP1 : UInt;
      State_Carrousel_P1TP2 : UInt;
      State_Carrousel_P3TP4 : UInt;
      State_Carrousel_P4TO : UInt;
      State_Carrousel : UInt;
   END_VAR
   VAR_TEMP
      i : UInt;
      j : UInt;
      f : UInt;
   END_VAR
BEGIN

   REGION TODO
       (*
       1. Need to confirm how the mode control is going to work, does switching the VTD to auto force all conveyors to auto as well or do we do seperate checks
       2. Need to review the shuttle interlock procedure inside the VTD function block
       *)

   END_REGION

   IF "FirstScan" THEN
       "OPC_Enable" := TRUE;
   END_IF;

   REGION Mode Control
       (*
           Mode select is done via the HMI. Might add external mode select switches.

           Mode select mask:
           0: Disabled
           1: Manual
           2: Semi-Auto
           3: Auto
           4: Teach
           5: Maintenance
       *)

       // IF #Mode_Change <> #Mode_Current THEN
       //     //Disable all devices
       //     "Mode_Change_F"(Mode := #Mode_Change);
       // END_IF;
   END_REGION

   REGION Errors VTD STATE
       IF #State_VTD > 30 AND #State_VTD < 120 THEN
           IF #Source_Location_VTD.Device_Type = 10 OR #Destination_Location_VTD.Device_Type = 10 THEN
               IF "Control_DB".LCnv_Control[#Source_Location_VTD.Level].Error
                   OR
                   "Control_DB".LCnv_Control[#Destination_Location_VTD.Level].Error THEN
                   "Error_Word_1".%X3 := TRUE;
                   #State_VTD := 400;
               END_IF;
           END_IF;
           IF "Control_DB".ECnv_Control.Error THEN
               "Error_Word_1".%X4 := TRUE;
               #State_VTD := 400;
           END_IF;
           IF "VTD_FB_DB".I_State = 400 THEN
               "Error_Word_1".%X5 := TRUE;
               #State_VTD := 400;
           END_IF;

       END_IF;
   END_REGION

   // REGION Errors CAROUSEL STATE
   //     IF #State_Carrousel > 30 AND #State_Carrousel < 120 THEN
   //         IF #Source_Location_Carousel.Device_Type = 10 OR #Destination_Location_VTD.Device_Type = 10 THEN
   //             IF "Control_DB".LCnv_Control[#Source_Location_Carousel.Level].Error
   //                 OR
   //                 "Control_DB".LCnv_Control[#Destination_Location_VTD.Level].Error THEN
   //                 #State_Carrousel := 400;
   //             END_IF;
   //         ELSIF #Source_Location_Carousel.Device_Type = 11 OR #Destination_Location_VTD.Device_Type = 11 THEN
   //             IF "Control_DB".LCnv_Control[#Source_Location_Carousel.Level].Error
   //                 OR
   //                 "Control_DB".LCnv_Control[#Destination_Location_VTD.Level].Error
   //             THEN
   //                 #State_Carrousel := 400;
   //             END_IF;
   //         END_IF;
   //         IF "Control_DB".ECnv_Control.Error THEN
   //             #State_Carrousel := 400;
   //         END_IF;
   //         IF "VTD_FB_DB".I_State = 400 THEN
   //             #State_Carrousel := 400;
   //         END_IF;

   //     END_IF;
   // END_REGION

   //Bit OPC in Error
   IF #State_VTD = 400 OR #State_Carrousel_CTC = 400 OR #State_Carrousel_ITP1 = 400 OR #State_Carrousel_P1TP2 = 400
       OR #State_Carrousel_P3TP4 = 400 OR #State_Carrousel_P4TO = 400 OR #State_Carrousel_P4TPICK = 400
       OR #State_Carrousel_PICKTP1 = 400
   THEN
       "Error_Word_1".%X0 := TRUE;
   ELSE
       "Error_Word_1".%X0 := FALSE;
   END_IF;

   REGION OPC UA Control
       (*
       Type of task to be performed:
           1 = Move to Floor
           2 = Shuttle Transfer into VTD
           3 = Shuttle Transfer out of VTD
           4 = Transfer Pallet into VTD
           5 = Transfer Pallet out of VTD
           6 = Transfer Pallet Roller to Roller
           7 = Transfer Pallet Chain to Chain  
           8 = Transfer to pick station 
           9 = Transfer from Pick station 
           10 = Weigh Pallet
           11 = Set chain Cnv as active (lower) // no use for now
           12 = Set Roller Cnv as active (raise) // no use for now

           Need to isolate ZZ in XXYYZZ to confirm #i = ZZ

           Extract XX (first two digits)
           xx := inputNumber / 10000;

           Extract YY (middle two digits)
           yy := (inputNumber / 100) MOD 100;

           Extract ZZ (last two digits)
           zz := inputNumber MOD 100;    
       *)

       REGION VTDs and Buffer conveyors
           IF "VTD_Buffers_In_Automatic" AND #OPC_Enable THEN
               CASE #State_VTD OF
                   0:  //Pre operational state
                       #State_VTD := 10;

                   10: //Idle waiting for task
                       IF "Control_DB"."VTD_Order Table".Task_Data_Available AND "Control_DB".VTD_Control.Mode = 3 AND
                           NOT "Control_DB".VTD_Control.Running AND NOT "Control_DB"."VTD_Order Table".Movement_Ready AND "Control_DB".VTD_Control.SM_State <= 10 THEN
                               // "Control_DB".WMS_OPC_UA.Task_Data_Available := FALSE;
                               #State_VTD := 20;
                           END_IF;

                   20: //Determine the type of task
                       "ID_Decode_F"(ID := "Control_DB"."VTD_Order Table".Source_Location,
                                     ID_Decoded := #Source_Location_VTD);
                       "ID_Decode_F"(ID := "Control_DB"."VTD_Order Table".Destination_Location,
                                     ID_Decoded := #Destination_Location_VTD);

                       //VTD move to floor
                       IF "Control_DB"."VTD_Order Table".Task_Type = 1
                           AND NOT "Control_DB".VTD_Control.Running THEN
                           #State_VTD := 30;

                           //Shuttle transfer in/out of the VTD
                       ELSIF "Control_DB"."VTD_Order Table".Task_Type = 2 OR "Control_DB"."VTD_Order Table".Task_Type = 3
                       THEN
                           #State_VTD := 70;

                           //Transfer Pallet in/out of the VTD
                       ELSIF "Control_DB"."VTD_Order Table".Task_Type = 4 OR "Control_DB"."VTD_Order Table".Task_Type = 5
                       THEN
                           #State_VTD := 100;
                       END_IF;

                           //=========================== VTD Move to floor ===========================
                       30: //Set all the Move to level variables
                           "Control_DB".VTD_Control.Current_Task_Type := INT_TO_UINT("Control_DB"."VTD_Order Table".Task_Type);
                           "Control_DB".VTD_Control.Instruction.Pallet_Type := "Control_DB"."VTD_Order Table".Pallet_Type;
                           "Control_DB".VTD_Control.Instruction.Task_ID := INT_TO_UINT("Control_DB"."VTD_Order Table".Task_ID);
                           "Control_DB".VTD_Control.Instruction.Task_Metadata := "Control_DB"."VTD_Order Table".Task_Metadata;
                           "Control_DB".VTD_Control.Instruction.Move_To_Level := INT_TO_UINT(#Destination_Location_VTD.Level);
                           #State_VTD := 35;

                       35://Wait for the VTD to start its movement
                           "Control_DB"."VTD_Order Table".SM_State := "Control_DB".VTD_Control.SM_State;
                           IF "Control_DB".VTD_Control.Enabled AND "Control_DB".VTD_Control.Running THEN
                               "Control_DB"."VTD_Order Table".Movement_Ready := TRUE;
                              // "Control_DB"."VTD_Order Table".Task_Data_Available := FALSE;//
                               #State_VTD := 40;
                           END_IF;

                       40: //Wait for the VTD to complete its movement
                           "Control_DB"."VTD_Order Table".SM_State := "Control_DB".VTD_Control.SM_State;
                           IF "Control_DB".VTD_Control.SM_State = 100 THEN

                               #State_VTD := 41;
                           END_IF;

                       41: //Wait for XXs for report done
                           "IEC_Timer_0_DB_6".TON(IN := TRUE,
                                                   PT := T#2000ms);
                            IF "IEC_Timer_0_DB_6".Q THEN
                                "Control_DB"."VTD_Order Table".Movement_Request_Complete := TRUE;
                                #State_VTD := 45;
                           END_IF;

                       45: //Wait for the ACK before we go back to Idle
                           "Control_DB"."VTD_Order Table".SM_State := "Control_DB".VTD_Control.SM_State;
                           IF "Control_DB"."VTD_Order Table".Movement_Request_Complete_Ack THEN///////////////////////////////////////////////////////////////////
                               // "Control_DB".WMS_OPC_UA.Task_Type := 0;
                               // "Control_DB".VTD_Control.Instruction.Reset := TRUE;///////////////////////////////////////////////////////////////////
                               #State_VTD := 250;
                           END_IF;

                           //=========================== Transfer Shuttle in/out of the VTD ===========================

                       70: //Set all the shuttle interlock variables
                           "Control_DB".VTD_Control.Instruction.Task_ID := "Control_DB"."VTD_Order Table".Task_ID; //Assign task ID to WCS Task ID
                           "Control_DB".VTD_Control.Instruction.Task_Metadata := "Control_DB"."VTD_Order Table".Task_Metadata;
                           "Control_DB".VTD_Control.Instruction.Pallet_Type := "Control_DB"."VTD_Order Table".Pallet_Type;
                           "Control_DB".VTD_Control.Current_Task_Type := INT_TO_UINT("Control_DB"."VTD_Order Table".Task_Type);
                           "Control_DB".VTD_Control.Shuttle_Interlock.Shuttle_Interlock_Task_ID := INT_TO_UINT("Control_DB"."VTD_Order Table".Task_ID);
                           "Control_DB".VTD_Control.Shuttle_Interlock.Shuttle_Interlock_Task_Metadata := "Control_DB"."VTD_Order Table".Task_Metadata;
                           "Control_DB".VTD_Control.Shuttle_Interlock.Shuttle_ID := INT_TO_UINT("Control_DB"."VTD_Order Table".Shuttle_ID);
                           "Control_DB".VTD_Control.Shuttle_Interlock.Shuttle_Loaded := "Control_DB"."VTD_Order Table".Shuttle_Loaded;
                           "Control_DB".VTD_Control.Shuttle_Interlock.Shuttle_Start_Location := "Control_DB"."VTD_Order Table".Source_Location;
                           "Control_DB".VTD_Control.Shuttle_Interlock.Shuttle_Target_Location := "Control_DB"."VTD_Order Table".Destination_Location;

                           "Control_DB".VTD_Control.Shuttle_Interlock.Interlock_Request := TRUE;
                           #State_VTD := 75;

                       75: //Inform WCS that the VTD is ready to interlock
                           "Control_DB"."VTD_Order Table".SM_State := "Control_DB".VTD_Control.SM_State;
                           IF "Control_DB".VTD_Control.Shuttle_Interlock.Ready_To_Interlock THEN
                               "Control_DB"."VTD_Order Table".Movement_Ready := TRUE;
                               "Control_DB"."VTD_Order Table".Task_Data_Available := FALSE;
                               #State_VTD := 80;
                           END_IF;

                       80://Inform WCS that the interlock is complete
                           IF "Control_DB".VTD_Control.Shuttle_Interlock.Interlock_Complete THEN
                               "Control_DB".VTD_Control.Shuttle_Interlock.Interlock_Request := FALSE;
                               "Control_DB"."VTD_Order Table".Movement_Request_Complete := TRUE;
                               #State_VTD := 81;
                           END_IF;

                       81: //Wait for XXs for report done
                           "IEC_Timer_0_DB_7".TON(IN := TRUE,
                                                   PT := T#500mS);
                           IF "IEC_Timer_0_DB_7".Q THEN
                               #State_VTD := 90;
                           END_IF;

                       90: //Reset VTD back to idle state
                           IF "Control_DB"."VTD_Order Table".Movement_Request_Complete_Ack THEN
                               "Control_DB".VTD_Control.Shuttle_Interlock.Interlock_Complete_Ack := TRUE;
                               #State_VTD := 250;
                           END_IF;

                           //=========================== Transfer Pallet in/out of the VTD ===========================

                       100: //Set the destination conveyor variables

                           //Assign task to receiving conveyor
                           IF #Destination_Location_VTD.Level >= "Settings_DB".VTD_Settings.Lowest_Level AND #Destination_Location_VTD.Level <= "Settings_DB".VTD_Settings.Highest_Level THEN

